       // Shuttle in Place Cnv_Inputs - Need to confirm the order of these Cnv_Inputs.
       // IF (#Cnv_Settings.ID > 110000 AND #Cnv_Settings.ID < 120000 AND NOT #Cnv_Control.Inputs.Sdetect1 AND #Cnv_Control.Inputs.Sdetect2)
       //     OR (#Cnv_Settings.ID > 120000 AND #Cnv_Settings.ID < 130000 AND NOT #Cnv_Control.Inputs.Sdetect1 AND #Cnv_Control.Inputs.Sdetect2) THEN
       //     #Cnv_Control.Error := TRUE; //14:5 Shuttle is about to yeet itself down the VTD shaft
       //     "Set_Bit_F"(Bit := 7,
       //                 Bit_Value := 1,
       //                 Var := #Cnv_Control.Cnv_Errors.Error_Word_2);
       //     #State := 400;
       // END_IF;

       // IF (#Cnv_Settings.ID > 110000 AND #Cnv_Settings.ID < 120000 AND #Cnv_Control.Inputs.Sdetect1 AND NOT #Cnv_Control.Inputs.Sdetect2)
       //     OR (#Cnv_Settings.ID > 120000 AND #Cnv_Settings.ID < 130000 AND #Cnv_Control.Inputs.Sdetect1 AND NOT #Cnv_Control.Inputs.Sdetect2) THEN
       //     #Cnv_Control.Warning := 0; //Shuttle detected in conveyor not yet on barcode
       // END_IF;

       // // #Watchdog auto starts the moment Any form OF transfer occurs.
       // IF #State > 10 AND #State < 400 THEN
       //     #Watchdog(IN := TRUE,
       //               PT := T#200s);
       // ELSE
       //     #Watchdog.IN := FALSE;
       // END_IF;

       // IF #Watchdog.Q THEN
       //     #Watchdog.IN := FALSE;
       //     #Cnv_Control.Error := TRUE; //14:2  Watchdog bit
       //     "Set_Bit_F"(Bit := 4,
       //                 Bit_Value := 1,
       //                 Var := #Cnv_Control.Cnv_Errors.Error_Word_2);
       //     #State := 400;
       // END_IF;

       // go to error state
       IF #Cnv_Control.Cnv_Errors.Error_Word_1 <> 0 OR
           #Cnv_Control.Cnv_Errors.Error_Word_2 <> 0 OR
           #Cnv_Control.Cnv_Errors.Error_Word_3 <> 0 OR
           #Cnv_Control.Cnv_Errors.Error_Word_4 <> 0
       THEN
           #Cnv_Control.Error := TRUE;
           #State := 400;
       END_IF;
   END_REGION

   REGION VFD
       REGION ROLLER
           #Cnv_Control.Roller_Motor.Ready := NOT #Cnv_Control.Roller_Motor.Error;

           #SinaSpeed_Roller(EnableAxis := #Cnv_Control.Roller_Motor.Forward OR #Cnv_Control.Roller_Motor.Reverse,
                             AckError := #Cnv_Control.Instruction.Reset,
                             SpeedSp := #MainSetpoint_Roller,
                             RefSpeed := 1745.0,
                             HWIDSTW := #Cnv_Settings.Roller_G120_Hardware_ID,
                             HWIDZSW := #Cnv_Settings.Roller_G120_Hardware_ID,
                             AxisEnabled => #Cnv_Control.Roller_Motor.Status.%X0,
                             Lockout => #Cnv_Control.Roller_Motor.Error,
                             Error => #Cnv_Control.Roller_Motor.Error);

           //MAIN SETPOINT
           IF #Cnv_Control.Roller_Motor.Reverse THEN
               #MainSetpoint_Roller := (SCALE_X(MIN := 0,
                                                VALUE := NORM_X(MIN := 0,
                                                                VALUE := #Cnv_Control.Roller_Motor.Speed,
                                                                MAX := 100),
                                                MAX := 1745.0) * -1);
           ELSIF #Cnv_Control.Roller_Motor.Forward THEN
               #MainSetpoint_Roller := SCALE_X(MIN := 0,
                                               VALUE := NORM_X(MIN := 0,
                                                               VALUE := #Cnv_Control.Roller_Motor.Speed,
                                                               MAX := 100),
                                               MAX := 1745.0);
           ELSE
               #MainSetpoint_Roller := 0;
           END_IF;

           REGION Actual Speed
               IF #MainSetpoint_Roller > 0 THEN
                   #Cnv_Control.Roller_Motor.Speed_Actual := SCALE_X(MIN := 0,
                                                                     VALUE := NORM_X(MIN := 0,
                                                                                     VALUE := #SinaSpeed_Roller.ActVelocity,
                                                                                     MAX := 1745.0),
                                                                     MAX := 100);
               ELSIF #MainSetpoint_Roller < 0 THEN
                   #Cnv_Control.Roller_Motor.Speed_Actual := SCALE_X(MIN := 0,
                                                                     VALUE := NORM_X(MIN := 0,
                                                                                     VALUE := #SinaSpeed_Roller.ActVelocity * -1,
                                                                                     MAX := 1745.0),
                                                                     MAX := 100);
               ELSE
                   #Cnv_Control.Roller_Motor.Speed_Actual := 0;
               END_IF;
           END_REGION
       END_REGION

       REGION CHAIN
           #Cnv_Control.Chain_Motor.Ready := NOT #Cnv_Control.Chain_Motor.Error;

           #SinaSpeed_Chain(EnableAxis := #Cnv_Control.Chain_Motor.Forward OR #Cnv_Control.Chain_Motor.Reverse,
                            AckError := #Cnv_Control.Instruction.Reset,
                            SpeedSp := #MainSetpoint_Chain,
                            RefSpeed := 1745.0,
                            HWIDSTW := #Cnv_Settings.Chain_G120_Hardware_ID,
                            HWIDZSW := #Cnv_Settings.Chain_G120_Hardware_ID,
                            AxisEnabled => #Cnv_Control.Chain_Motor.Status.%X0,
                            Lockout => #Cnv_Control.Chain_Motor.Error,
                            Error => #Cnv_Control.Chain_Motor.Error);

           //MAIN SETPOINT
           IF #Cnv_Control.Chain_Motor.Reverse THEN
               #MainSetpoint_Chain := (SCALE_X(MIN := 0,
                                               VALUE := NORM_X(MIN := 0,
                                                               VALUE := #Cnv_Control.Chain_Motor.Speed,
                                                               MAX := 100),
                                               MAX := 1745.0) * -1);
           ELSIF #Cnv_Control.Chain_Motor.Forward THEN
               #MainSetpoint_Chain := SCALE_X(MIN := 0,
                                              VALUE := NORM_X(MIN := 0,
                                                              VALUE := #Cnv_Control.Chain_Motor.Speed,
                                                              MAX := 100),
                                              MAX := 1745.0);
           ELSE
               #MainSetpoint_Chain := 0;
           END_IF;

           REGION Actual Speed
               IF #MainSetpoint_Chain > 0 THEN
                   #Cnv_Control.Chain_Motor.Speed_Actual := SCALE_X(MIN := 0,
                                                                    VALUE := NORM_X(MIN := 0,
                                                                                    VALUE := #SinaSpeed_Chain.ActVelocity,
                                                                                    MAX := 1745.0),
                                                                    MAX := 100);
               ELSIF #MainSetpoint_Chain < 0 THEN
                   #Cnv_Control.Chain_Motor.Speed_Actual := SCALE_X(MIN := 0,
                                                                    VALUE := NORM_X(MIN := 0,
                                                                                    VALUE := #SinaSpeed_Chain.ActVelocity * -1,
                                                                                    MAX := 1745.0),
                                                                    MAX := 100);
               ELSE
                   #Cnv_Control.Chain_Motor.Speed_Actual := 0;
               END_IF;
           END_REGION
       END_REGION

       REGION LIFT
           #Cnv_Control.Lift_Motor.Ready := NOT #Cnv_Control.Lift_Motor.Error;

           #SinaSpeed_Lift(EnableAxis := #Cnv_Control.Lift_Motor.Forward OR #Cnv_Control.Lift_Motor.Reverse,
                           AckError := #Cnv_Control.Instruction.Reset,
                           SpeedSp := #MainSetpoint_Lift,
                           RefSpeed := 1745.0,
                           HWIDSTW := #Cnv_Settings.Lift_G120_Hardware_ID,
                           HWIDZSW := #Cnv_Settings.Lift_G120_Hardware_ID,
                           AxisEnabled => #Cnv_Control.Lift_Motor.Status.%X0,
                           Lockout => #Cnv_Control.Lift_Motor.Error,
                           Error => #Cnv_Control.Lift_Motor.Error);

           //MAIN SETPOINT
           IF #Cnv_Control.Lift_Motor.Reverse THEN
               #MainSetpoint_Lift := (SCALE_X(MIN := 0,
                                              VALUE := NORM_X(MIN := 0,
                                                              VALUE := #Cnv_Control.Lift_Motor.Speed,
                                                              MAX := 100),
                                              MAX := 1745.0) * -1);
           ELSIF #Cnv_Control.Lift_Motor.Forward THEN
               #MainSetpoint_Lift := SCALE_X(MIN := 0,
                                             VALUE := NORM_X(MIN := 0,
                                                             VALUE := #Cnv_Control.Lift_Motor.Speed,
                                                             MAX := 100),
                                             MAX := 1745.0);
           ELSE
               #MainSetpoint_Lift := 0;
           END_IF;

           REGION Actual Speed
               IF #MainSetpoint_Lift > 0 THEN
                   #Cnv_Control.Lift_Motor.Speed_Actual := SCALE_X(MIN := 0,
                                                                   VALUE := NORM_X(MIN := 0,
                                                                                   VALUE := #SinaSpeed_Lift.ActVelocity,
                                                                                   MAX := 1745.0),
                                                                   MAX := 100);
               ELSIF #MainSetpoint_Lift < 0 THEN
                   #Cnv_Control.Lift_Motor.Speed_Actual := SCALE_X(MIN := 0,
                                                                   VALUE := NORM_X(MIN := 0,
                                                                                   VALUE := #SinaSpeed_Lift.ActVelocity * -1,
                                                                                   MAX := 1745.0),
                                                                   MAX := 100);
               ELSE
                   #Cnv_Control.Lift_Motor.Speed_Actual := 0;
               END_IF;
           END_REGION
       END_REGION
   END_REGION
END_FUNCTION_BLOCK

FUNCTION_BLOCK "PConveyor_4_FB"   // FB27, SCL
TITLE = Conveyor Instance FB
{ S7_Optimized_Access := 'TRUE' }
AUTHOR : Mertin Coetzee
VERSION : 0.1
// stored: AutoNumber true, IsIECCheckEnabled false, IsRetainMemResEnabled false, MemoryReserve 100, SetENOAutomatically false, UDAEnableTagReadback false
   VAR_INPUT
      Cnv_Settings : "PopUp_Cnv_Settings";
      TimeStartBoost_Roller : UInt;
   END_VAR
   VAR_IN_OUT
      Cnv_Control : "PopUp_Cnv_Control";
      SinaSpeed_Roller : SinaSpeed;
      SinaSpeed_Lift : SinaSpeed;
   END_VAR
   VAR
      State : UInt;
      Timer_TC : TON_TIME;
      Timer_Transfer { S7_SetPoint := 'True'} : TON_TIME;
      Watchdog { S7_SetPoint := 'True'} : TON_TIME;
      Transfer_Direction { S7_SetPoint := 'True'} : String;
      MainSetpoint_Roller : Int;
      MainSetpoint_Lift : Int;
      IEC_Timer_0_Instance_1 { S7_SetPoint := 'True'} : TON_TIME;
      R_TRIG_Instance { S7_SetPoint := 'True'} : R_TRIG;
   END_VAR
   VAR_TEMP
      Execute_Old : Bool;
      Stop_Old : Bool;
   END_VAR
BEGIN
   "R_TRIG_DB_23"(CLK := #Cnv_Control.Instruction.Execute AND NOT #Execute_Old);
   "R_TRIG_DB_24"(CLK := #Cnv_Control.Instruction.Stop AND NOT #Stop_Old);

   #Execute_Old := #Cnv_Control.Instruction.Execute;
   #Stop_Old := #Cnv_Control.Instruction.Stop;

   #Cnv_Control.Enabled := #Cnv_Control.Instruction.Enable;

   //MODES
   #Cnv_Control.Mode := #Cnv_Control.Instruction.Mode_Change;
   IF (#Cnv_Control.Mode = 1 OR #Cnv_Control.Mode = 5) AND NOT #Cnv_Control.Error THEN
       #State := 500;
   END_IF;

   #R_TRIG_Instance(CLK := #Cnv_Control.Mode = 3);
   IF #R_TRIG_Instance.Q THEN
       #State := 0;
   END_IF;

   (*
   TODO:
   01. Need to add statemachine watchdog - Done
   02. Extractor needs to be on same floor for pallet to be moved in manual passed Rbwd - Done
   03. Complete reset state - Done
   04. Add stop inputs - Done
   05. Need to add variable motor speed, manual needs to be slower. - Done
   06. Need to add cyclic error checking. For odd sensor combinations as well - Partially done
   07. Need to add Shuttle monitor - Done
   08. Need to add Task ID check and start bit check to outbound pallet move. Check direction of pallet movement based on connected Cnv.
   09. Need to add checks for wrong direction of travel - Done
   10. Add checks for unsafe conditions with Cnv_Inputs - Partially Done
   11. Define Error codes - DOne
   12. Add watchdof time to Cnv Settings - Done
   13. Add self-timeout on manual 
   14. For shuttle in place sensor checks take into account extractor floor and safety stopper state
   15. Confirm modes and states are correct (Semi-auto and maintenance as well)
   16. Add the correct transfer process for the logistex-spacemaker pallet handovers.

   Mode select is done via the HMI. Might add external mode select switches.

           Mode select mask:
           0: Disabled
           1: Manual
           2: Semi-Auto
           3: Auto
           4: Teach - N/A for Cnv
           5: Maintenance

   Device ID Format: XXYYZZ    
   XX = Device type   
       01   VTD
       10  Cnv_Front_of_VTD
       11  Cnv_Rear_of_VTD
       12  Cnv_On_Extractor
       20  Safety_Stop_Front_of_VTD
       21  Safety_Stop_Rear_of_VTD
   YY = Floor   
   ZZ = VTD Connected to    
   Example: 110203 Conveyor at the rear of VTD 3 on level 2

   Pallet Alignment
   0 = no alignment
   1 = center alignment
   2 = Left
   3 = Right

    Sensor order for the conveyor:
    Lfwd Lpd1 Lpd2
     []   []   []
    ##############################
    #        Pallet Flow         #
    #         ------->>          #
    #                            #
    #                            #
    ##############################
                     []   []   []
                    Rpd2 Rpd1 Rbwd      
   *)


   REGION Cyclic Checks    
       #Cnv_Control.Cnv_Occupied := "PopUp Conveyor 4 - Pallet present 1";

       // Update the Cnv_Control opbject
       #Cnv_Control.SM_State := #State;
       #Cnv_Control.Stopped := NOT #Cnv_Control.Running;
       IF #Cnv_Control.Instruction.Inbound_Ready OR #Cnv_Control.Instruction.Outbound_Ready THEN
           #Cnv_Control.Ready_For_Task := TRUE;
       ELSE
           #Cnv_Control.Ready_For_Task := FALSE;
       END_IF;

   END_REGION

   REGION Auto/Semi auto mode
       CASE #State OF
           0: //IDLE MODE
               #Cnv_Control.Instruction.Transfer_Complete := 0;
               #Cnv_Control.Instruction.Transfer_in_Progress := FALSE;
               #Cnv_Control.Running := FALSE;
               #Cnv_Control.Running := FALSE;
               #Cnv_Control.Roller_Motor.Forward := FALSE;
               #Cnv_Control.Roller_Motor.Reverse := FALSE;
               #Cnv_Control.Roller_Motor.Speed := 0;
               #Cnv_Control.Chain_Motor.Forward := FALSE;
               #Cnv_Control.Chain_Motor.Reverse := FALSE;
               #Cnv_Control.Chain_Motor.Speed := 0;
               #Cnv_Control.Lift_Motor.Forward := FALSE;
               #Cnv_Control.Lift_Motor.Reverse := FALSE;
               #Cnv_Control.Lift_Motor.Speed := 0;
               #Transfer_Direction := '';
               #Timer_Transfer(IN := FALSE,
                               PT := T#0ms);
               "IEC_Timer_0_DB_25".TON(IN := FALSE,
                                       PT := t#0s);
               IF #Cnv_Control.Enabled AND (#Cnv_Control.Mode = 3 OR #Cnv_Control.Mode = 2) AND #Cnv_Control.Error = 0 THEN
                   #State := 10;
               END_IF;

           10: //Standby - Conveyor ready to receive instruction
               IF ("R_TRIG_DB_23".Q OR #Cnv_Control.Instruction.Start_Transfer) THEN
                   //Inbound Transfer
                   IF #Cnv_Control.Instruction.Inbound_Ready AND NOT #Cnv_Control.Running AND #Cnv_Control.Error = 0 THEN
                       IF #Cnv_Control.Inputs."Lift Up" THEN
                           #Cnv_Control.Done := FALSE;
                           #Cnv_Control.Instruction.Transfer_in_Progress := TRUE;
                           #Cnv_Control.Current_Task_ID := #Cnv_Control.Instruction.Task_ID;
                           #State := 20;
                       END_IF;
                       //Outbound Transfer    
                   ELSIF #Cnv_Control.Instruction.Outbound_Ready AND NOT #Cnv_Control.Running AND #Cnv_Control.Error = 0 THEN
                       IF #Cnv_Control.Inputs."Lift Up" THEN
                           #Cnv_Control.Done := FALSE;
                           #Cnv_Control.Instruction.Transfer_in_Progress := TRUE;
                           #Cnv_Control.Current_Task_ID := #Cnv_Control.Instruction.Task_ID;
                           #State := 30;
                       END_IF;
                   END_IF;
               END_IF;

               IF #Cnv_Control.Instruction.Lift_Up THEN
                   #Cnv_Control.Done := FALSE;
                   #State := 60; // Lift UP
               ELSIF #Cnv_Control.Instruction.Lift_Down THEN
                   #Cnv_Control.Done := FALSE;
                   #State := 70; // Lift Down
               END_IF;

           20: // Roller Running (Popup Up)
               #Cnv_Control.Running := TRUE;
               #Cnv_Control.Roller_Motor.Forward := TRUE;
               "IEC_Timer_0_DB_25".TON(IN := TRUE,
                                       PT := UINT_TO_TIME(#TimeStartBoost_Roller) * 1000);

               IF NOT "IEC_Timer_0_DB_25".Q THEN
                   #Cnv_Control.Roller_Motor.Speed := 100.0;
               ELSE
                   #Cnv_Control.Roller_Motor.Speed := #Cnv_Settings.Roller_Full_Speed;
               END_IF;

               #Transfer_Direction := 'Foward';

               IF "R_TRIG_DB_24".Q OR "PopUp Conveyor 4 - Pallet present 1" THEN
                   "IEC_Timer_0_DB_25".TON(IN := FALSE,
                                           PT := t#0s);
                   #Cnv_Control.Done := TRUE;
                   #Cnv_Control.Roller_Motor.Forward := FALSE;
                   #Cnv_Control.Roller_Motor.Reverse := FALSE;
                   #Cnv_Control.Roller_Motor.Speed := 0;
                   #Transfer_Direction := '';
                   #State := 0;
               END_IF;

               //Monitor the transfer progress
               #Timer_Transfer(IN := TRUE,
                               PT := UINT_TO_TIME(#Cnv_Settings.Roller_Transfer_Time) * 1000);
               //If the watchdog bites, kill the process
               IF #Timer_Transfer.Q THEN //14:1 Transfer timed out
                   "Set_Bit_F"(Bit := 3,
                               Bit_Value := 1,
                               Var := #Cnv_Control.Cnv_Errors.Error_Word_2);
               END_IF;

           30: // Roller Running (Popup Up)
               IF "Control_DB".Outbound_Cnv.Motor.Status.%X0 THEN
                   #Cnv_Control.Running := TRUE;
                   #Cnv_Control.Roller_Motor.Forward := TRUE;
                   #Cnv_Control.Roller_Motor.Speed := #Cnv_Settings.Roller_Full_Speed;
                   #Transfer_Direction := 'Foward';
               END_IF;

               IF "R_TRIG_DB_24".Q OR NOT "Outbound Conveyor" THEN
                   #Cnv_Control.Done := TRUE;
                   #Cnv_Control.Roller_Motor.Forward := FALSE;
                   #Cnv_Control.Roller_Motor.Reverse := FALSE;
                   #Cnv_Control.Roller_Motor.Speed := 0;
                   #Transfer_Direction := '';
                   #State := 0;
               END_IF;

               //Monitor the transfer progress
               #Timer_Transfer(IN := TRUE,
                               PT := UINT_TO_TIME(#Cnv_Settings.Roller_Transfer_Time) * 1000);
               //If the watchdog bites, kill the process
               IF #Timer_Transfer.Q THEN //14:1 Transfer timed out
                   "Set_Bit_F"(Bit := 3,
                               Bit_Value := 1,
                               Var := #Cnv_Control.Cnv_Errors.Error_Word_2);
               END_IF;

           60: // Lift Up
               #Cnv_Control.Running := TRUE;
               #Cnv_Control.Lift_Motor.Forward := TRUE;
               #Cnv_Control.Lift_Motor.Speed := #Cnv_Settings.Lift_Full_Speed;
               #Transfer_Direction := 'Up';

               IF #Cnv_Control.Inputs."Lift Up" THEN
                   #Cnv_Control.Done := TRUE;
                   #Cnv_Control.Lift_Motor.Forward := FALSE;
                   #Cnv_Control.Lift_Motor.Reverse := FALSE;
                   #Cnv_Control.Lift_Motor.Speed := 0;
                   #Transfer_Direction := '';
                   #State := 0;
               END_IF;

               //Monitor the transfer progress
               #Timer_Transfer(IN := TRUE,
                               PT := UINT_TO_TIME(#Cnv_Settings.Lift_Transfer_Time) * 1000);
               //If the watchdog bites, kill the process
               IF #Timer_Transfer.Q THEN //14:1 Transfer timed out
                   "Set_Bit_F"(Bit := 3,
                               Bit_Value := 1,
                               Var := #Cnv_Control.Cnv_Errors.Error_Word_2);
               END_IF;

           70: // Lift Down
               #Cnv_Control.Running := TRUE;
               #Cnv_Control.Lift_Motor.Reverse := TRUE;
               #Cnv_Control.Lift_Motor.Speed := #Cnv_Settings.Lift_Full_Speed;
               #Transfer_Direction := 'Down';

               IF #Cnv_Control.Inputs."Lift Down" THEN
                   #Cnv_Control.Done := TRUE;
                   #Cnv_Control.Lift_Motor.Forward := FALSE;
                   #Cnv_Control.Lift_Motor.Reverse := FALSE;
                   #Cnv_Control.Lift_Motor.Speed := 0;
                   #Transfer_Direction := '';
                   #State := 0;
               END_IF;

               //Monitor the transfer progress
               #Timer_Transfer(IN := TRUE,
                               PT := UINT_TO_TIME(#Cnv_Settings.Lift_Transfer_Time) * 1000);
               //If the watchdog bites, kill the process
               IF #Timer_Transfer.Q THEN //14:1 Transfer timed out
                   "Set_Bit_F"(Bit := 3,
                               Bit_Value := 1,
                               Var := #Cnv_Control.Cnv_Errors.Error_Word_2);
               END_IF;

           400: //Error state
               #Cnv_Control.Running := FALSE;
               #Cnv_Control.Roller_Motor.Speed := 0;
               #Cnv_Control.Chain_Motor.Speed := 0;
               #Cnv_Control.Lift_Motor.Speed := 0;
               #Cnv_Control.Roller_Motor.Forward := FALSE;
               #Cnv_Control.Chain_Motor.Forward := FALSE;
               #Cnv_Control.Lift_Motor.Forward := FALSE;
               #Cnv_Control.Roller_Motor.Reverse := FALSE;
               #Cnv_Control.Chain_Motor.Reverse := FALSE;
               #Cnv_Control.Lift_Motor.Reverse := FALSE;
               #Cnv_Control.Instruction.Stop := FALSE;
               #Cnv_Control.Instruction.Transfer_in_Progress := FALSE;
               #Watchdog(IN := FALSE,
                         PT := T#0S);
               #Timer_TC(IN := FALSE,
                         PT := T#0S);
               #Timer_Transfer(IN := FALSE,
                               PT := T#0S);
               #IEC_Timer_0_Instance_1(IN := FALSE,
                                       PT := T#0S);
               IF #Cnv_Control.Instruction.Reset THEN
                   #Cnv_Control.Warning := 0;
                   #Cnv_Control.Current_Task_ID := 0;
                   #Cnv_Control.Error := FALSE; //Reset the conveyor

                   #Cnv_Control.Cnv_Errors.Error_Word_1 := 0;
                   #Cnv_Control.Cnv_Errors.Error_Word_2 := 0;
                   #Cnv_Control.Cnv_Errors.Error_Word_3 := 0;
                   #Cnv_Control.Cnv_Errors.Error_Word_4 := 0;
                   #State := 0;
               END_IF;

           500:
               IF #Cnv_Control.Enabled THEN
                   REGION ROLLER
                       IF #Cnv_Control.Inputs."Lift Up" AND NOT #Cnv_Control.Inputs."Lift Down" THEN
                           IF #Cnv_Control.Instruction.Roller_Fwd OR #Cnv_Control.Instruction.Start_Transfer THEN
                               #Cnv_Control.Roller_Motor.Speed := #Cnv_Settings.Roller_Manual_Speed;
                               #Cnv_Control.Roller_Motor.Forward := TRUE;
                               #Cnv_Control.Running := TRUE;
                           ELSIF #Cnv_Control.Instruction.Roller_Bwd OR #Cnv_Control.Instruction.Start_Transfer_Backward THEN
                               #Cnv_Control.Roller_Motor.Speed := #Cnv_Settings.Roller_Manual_Speed;
                               #Cnv_Control.Roller_Motor.Reverse := TRUE;
                               #Cnv_Control.Running := TRUE;
                           ELSE
                               #Cnv_Control.Roller_Motor.Speed := 0;
                               #Cnv_Control.Roller_Motor.Forward := FALSE;
                               #Cnv_Control.Roller_Motor.Reverse := FALSE;
                               #Cnv_Control.Running := FALSE;
                           END_IF;
                       END_IF;
                   END_REGION

                   REGION LIFT
                       IF NOT #SinaSpeed_Roller.AxisEnabled THEN
                           IF #Cnv_Control.Instruction.Lift_Up AND NOT #Cnv_Control.Inputs."Lift Up" THEN
                               #Cnv_Control.Lift_Motor.Speed := #Cnv_Settings.Lift_Manual_Speed;
                               #Cnv_Control.Lift_Motor.Forward := TRUE;
                               #Cnv_Control.Running := TRUE;
                           ELSIF #Cnv_Control.Instruction.Lift_Down AND NOT #Cnv_Control.Inputs."Lift Down" THEN
                               #Cnv_Control.Lift_Motor.Speed := #Cnv_Settings.Lift_Manual_Speed;
                               #Cnv_Control.Lift_Motor.Reverse := TRUE;
                               #Cnv_Control.Running := TRUE;
                           ELSE
                               #Cnv_Control.Lift_Motor.Speed := 0;
                               #Cnv_Control.Lift_Motor.Forward := FALSE;
                               #Cnv_Control.Lift_Motor.Reverse := FALSE;
                               #Cnv_Control.Running := FALSE;
                           END_IF;
                       END_IF;
                   END_REGION
               END_IF;

               IF #Cnv_Control.Mode <> 1 AND #Cnv_Control.Mode <> 5 THEN
                   #State := 0;
               END_IF;
       END_CASE;
   END_REGION



   REGION Cyclic Error Checks
       IF NOT "Main_Safety_RTG1_DB".SAFETY_OK_CAROUSEL THEN //11:1
           "Set_Bit_F"(Bit := 0,
                       Bit_Value := 1,
                       Var := #Cnv_Control.Cnv_Errors.Error_Word_1);
       END_IF;

       // IF #Cnv_Control.Instruction.Stop THEN //11:2
       //     "Set_Bit_F"(Bit := 1,
       //                 Bit_Value := 1,
       //                 Var := #Cnv_Control.Cnv_Errors.Error_Word_1);
       // END_IF;

       IF #Cnv_Control.Roller_Motor.Error OR #Cnv_Control.Chain_Motor.Error OR #Cnv_Control.Lift_Motor.Error THEN
           "Set_Bit_F"(Bit := 0,
                       Bit_Value := 1,
                       Var := #Cnv_Control.Cnv_Errors.Error_Word_4);
       END_IF;

       // Pallet Sensor Checks
       // IF #Cnv_Control.Inputs.Lfwd AND #Cnv_Control.Inputs.Rbwd THEN
       //     #Cnv_Control.Error := TRUE; //15:2 Combination of Cnv_Inputs indicates issue in conveyor
       //     "Set_Bit_F"(Bit := 1,
       //                 Bit_Value := 1,
       //                 Var := #Cnv_Control.Cnv_Errors.Error_Word_4);
       //     #State := 400;
       // IF #Cnv_Control.Inputs.Lfwd AND #Cnv_Control.Inputs.Lpd1 AND #Cnv_Control.Inputs.Rpd1 THEN
       //     #Cnv_Control.Error := TRUE; //15:3 Combination of Cnv_Inputs indicates issue in conveyor
       //     "Set_Bit_F"(Bit := 2,
       //                 Bit_Value := 1,
       //                 Var := #Cnv_Control.Cnv_Errors.Error_Word_4);
       //     #State := 400;
       // ELSIF #Cnv_Control.Inputs.Rbwd AND #Cnv_Control.Inputs.Lpd1 AND #Cnv_Control.Inputs.Rpd1 THEN
       //     #Cnv_Control.Error := TRUE; //15:4 Combination of Cnv_Inputs indicates issue in conveyor
       //     "Set_Bit_F"(Bit := 3,
       //                 Bit_Value := 1,
       //                 Var := #Cnv_Control.Cnv_Errors.Error_Word_4);
       //     #State := 400;
       // END_IF;

       // Shuttle in Place Cnv_Inputs - Need to confirm the order of these Cnv_Inputs.
       // IF (#Cnv_Settings.ID > 110000 AND #Cnv_Settings.ID < 120000 AND NOT #Cnv_Control.Inputs.Sdetect1 AND #Cnv_Control.Inputs.Sdetect2)
       //     OR (#Cnv_Settings.ID > 120000 AND #Cnv_Settings.ID < 130000 AND NOT #Cnv_Control.Inputs.Sdetect1 AND #Cnv_Control.Inputs.Sdetect2) THEN
       //     #Cnv_Control.Error := TRUE; //14:5 Shuttle is about to yeet itself down the VTD shaft
       //     "Set_Bit_F"(Bit := 7,
       //                 Bit_Value := 1,
       //                 Var := #Cnv_Control.Cnv_Errors.Error_Word_2);
       //     #State := 400;
       // END_IF;

       // IF (#Cnv_Settings.ID > 110000 AND #Cnv_Settings.ID < 120000 AND #Cnv_Control.Inputs.Sdetect1 AND NOT #Cnv_Control.Inputs.Sdetect2)
       //     OR (#Cnv_Settings.ID > 120000 AND #Cnv_Settings.ID < 130000 AND #Cnv_Control.Inputs.Sdetect1 AND NOT #Cnv_Control.Inputs.Sdetect2) THEN
       //     #Cnv_Control.Warning := 0; //Shuttle detected in conveyor not yet on barcode
       // END_IF;

       // // #Watchdog auto starts the moment Any form OF transfer occurs.
       // IF #State > 10 AND #State < 400 THEN
       //     #Watchdog(IN := TRUE,
       //               PT := T#200s);
       // ELSE
       //     #Watchdog.IN := FALSE;
       // END_IF;

       // IF #Watchdog.Q THEN
       //     #Watchdog.IN := FALSE;
       //     #Cnv_Control.Error := TRUE; //14:2  Watchdog bit
       //     "Set_Bit_F"(Bit := 4,
       //                 Bit_Value := 1,
       //                 Var := #Cnv_Control.Cnv_Errors.Error_Word_2);
       //     #State := 400;
       // END_IF;

       // go to error state
       IF #Cnv_Control.Cnv_Errors.Error_Word_1 <> 0 OR
           #Cnv_Control.Cnv_Errors.Error_Word_2 <> 0 OR
           #Cnv_Control.Cnv_Errors.Error_Word_3 <> 0 OR
           #Cnv_Control.Cnv_Errors.Error_Word_4 <> 0
       THEN
           #Cnv_Control.Error := TRUE;
           #State := 400;
       END_IF;
   END_REGION

   REGION VFD
       REGION ROLLER
           #Cnv_Control.Roller_Motor.Ready := NOT #Cnv_Control.Roller_Motor.Error;

           #SinaSpeed_Roller(EnableAxis := #Cnv_Control.Roller_Motor.Forward OR #Cnv_Control.Roller_Motor.Reverse,
                             AckError := #Cnv_Control.Instruction.Reset,
                             SpeedSp := #MainSetpoint_Roller,
                             RefSpeed := 1745.0,
                             HWIDSTW := #Cnv_Settings.Roller_G120_Hardware_ID,
                             HWIDZSW := #Cnv_Settings.Roller_G120_Hardware_ID,
                             AxisEnabled => #Cnv_Control.Roller_Motor.Status.%X0,
                             Lockout => #Cnv_Control.Roller_Motor.Error,
                             Error => #Cnv_Control.Roller_Motor.Error);

           //MAIN SETPOINT
           IF #Cnv_Control.Roller_Motor.Reverse THEN
               #MainSetpoint_Roller := (SCALE_X(MIN := 0,
                                                VALUE := NORM_X(MIN := 0,
                                                                VALUE := #Cnv_Control.Roller_Motor.Speed,
                                                                MAX := 100),
                                                MAX := 1745.0) * -1);
           ELSIF #Cnv_Control.Roller_Motor.Forward THEN
               #MainSetpoint_Roller := SCALE_X(MIN := 0,
                                               VALUE := NORM_X(MIN := 0,
                                                               VALUE := #Cnv_Control.Roller_Motor.Speed,
                                                               MAX := 100),
                                               MAX := 1745.0);
           ELSE
               #MainSetpoint_Roller := 0;
           END_IF;

           REGION Actual Speed
               IF #MainSetpoint_Roller > 0 THEN
                   #Cnv_Control.Roller_Motor.Speed_Actual := SCALE_X(MIN := 0,
                                                                     VALUE := NORM_X(MIN := 0,
                                                                                     VALUE := #SinaSpeed_Roller.ActVelocity,
                                                                                     MAX := 1745.0),
                                                                     MAX := 100);
               ELSIF #MainSetpoint_Roller < 0 THEN
                   #Cnv_Control.Roller_Motor.Speed_Actual := SCALE_X(MIN := 0,
                                                                     VALUE := NORM_X(MIN := 0,
                                                                                     VALUE := #SinaSpeed_Roller.ActVelocity * -1,
                                                                                     MAX := 1745.0),
                                                                     MAX := 100);
               ELSE
                   #Cnv_Control.Roller_Motor.Speed_Actual := 0;
               END_IF;
           END_REGION
       END_REGION

       REGION LIFT
           #Cnv_Control.Lift_Motor.Ready := NOT #Cnv_Control.Lift_Motor.Error;

           #SinaSpeed_Lift(EnableAxis := #Cnv_Control.Lift_Motor.Forward OR #Cnv_Control.Lift_Motor.Reverse,
                           AckError := #Cnv_Control.Instruction.Reset,
                           SpeedSp := #MainSetpoint_Lift,
                           RefSpeed := 1745.0,
                           HWIDSTW := #Cnv_Settings.Lift_G120_Hardware_ID,
                           HWIDZSW := #Cnv_Settings.Lift_G120_Hardware_ID,
                           AxisEnabled => #Cnv_Control.Lift_Motor.Status.%X0,
                           Lockout => #Cnv_Control.Lift_Motor.Error,
                           Error => #Cnv_Control.Lift_Motor.Error);

           //MAIN SETPOINT
           IF #Cnv_Control.Lift_Motor.Reverse THEN
               #MainSetpoint_Lift := (SCALE_X(MIN := 0,
                                              VALUE := NORM_X(MIN := 0,
                                                              VALUE := #Cnv_Control.Lift_Motor.Speed,
                                                              MAX := 100),
                                              MAX := 1745.0) * -1);
           ELSIF #Cnv_Control.Lift_Motor.Forward THEN
               #MainSetpoint_Lift := SCALE_X(MIN := 0,
                                             VALUE := NORM_X(MIN := 0,
                                                             VALUE := #Cnv_Control.Lift_Motor.Speed,
                                                             MAX := 100),
                                             MAX := 1745.0);
           ELSE
               #MainSetpoint_Lift := 0;
           END_IF;

           REGION Actual Speed
               IF #MainSetpoint_Lift > 0 THEN
                   #Cnv_Control.Lift_Motor.Speed_Actual := SCALE_X(MIN := 0,
                                                                   VALUE := NORM_X(MIN := 0,
                                                                                   VALUE := #SinaSpeed_Lift.ActVelocity,
                                                                                   MAX := 1745.0),
                                                                   MAX := 100);
               ELSIF #MainSetpoint_Lift < 0 THEN
                   #Cnv_Control.Lift_Motor.Speed_Actual := SCALE_X(MIN := 0,
                                                                   VALUE := NORM_X(MIN := 0,
                                                                                   VALUE := #SinaSpeed_Lift.ActVelocity * -1,
                                                                                   MAX := 1745.0),
                                                                   MAX := 100);
               ELSE
                   #Cnv_Control.Lift_Motor.Speed_Actual := 0;
               END_IF;
           END_REGION
       END_REGION
   END_REGION
END_FUNCTION_BLOCK

FUNCTION_BLOCK "PickConveyor_FB"   // FB35, SCL
TITLE = Conveyor Instance FB
{ S7_Optimized_Access := 'TRUE' }
AUTHOR : Mertin Coetzee
VERSION : 0.1
// stored: AutoNumber true, IsIECCheckEnabled false, IsRetainMemResEnabled false, MemoryReserve 100, SetENOAutomatically false, UDAEnableTagReadback false
   VAR_INPUT
      Cnv_Settings : "Pick_Cnv_Settings";
   END_VAR
   VAR_IN_OUT
      SinaSpeed_Chain : SinaSpeed;
   END_VAR
   VAR
      State : UInt;
      Timer_TC : TON_TIME;
      Timer_Transfer { S7_SetPoint := 'True'} : TON_TIME;
      Watchdog { S7_SetPoint := 'True'} : TON_TIME;
      Transfer_Direction { S7_SetPoint := 'True'} : String;
      MainSetpoint_Chain : Int;
      IEC_Timer_0_Instance_1 { S7_SetPoint := 'True'} : TON_TIME;
      R_TRIG_Instance { S7_SetPoint := 'True'} : R_TRIG;
   END_VAR
   VAR_TEMP
      Execute_Old : Bool;
      Stop_Old : Bool;
   END_VAR
BEGIN
   "R_TRIG_DB_28"(CLK := "Control_DB".Pick_Station.Instruction.Execute AND NOT #Execute_Old);
   "R_TRIG_DB_29"(CLK := "Control_DB".Pick_Station.Instruction.Stop AND NOT #Stop_Old);

   #Execute_Old := "Control_DB".Pick_Station.Instruction.Execute;
   #Stop_Old := "Control_DB".Pick_Station.Instruction.Stop;

   "Control_DB".Pick_Station.Enabled := "Control_DB".Pick_Station.Instruction.Enable;

   //MODES
   "Control_DB".Pick_Station.Mode := "Control_DB".Pick_Station.Instruction.Mode_Change;
   IF ("Control_DB".Pick_Station.Mode = 1 OR "Control_DB".Pick_Station.Mode = 5) AND NOT "Control_DB".Pick_Station.Error THEN
       #State := 500;
   END_IF;

   #R_TRIG_Instance(CLK := "Control_DB".Pick_Station.Mode = 3);
   IF #R_TRIG_Instance.Q THEN
       #State := 0;
   END_IF;

   (*
   TODO:
   01. Need to add statemachine watchdog - Done
   02. Extractor needs to be on same floor for pallet to be moved in manual passed Rbwd - Done
   03. Complete reset state - Done
   04. Add stop inputs - Done
   05. Need to add variable motor speed, manual needs to be slower. - Done
   06. Need to add cyclic error checking. For odd sensor combinations as well - Partially done
   07. Need to add Shuttle monitor - Done
   08. Need to add Task ID check and start bit check to outbound pallet move. Check direction of pallet movement based on connected Cnv.
   09. Need to add checks for wrong direction of travel - Done
   10. Add checks for unsafe conditions with Cnv_Inputs - Partially Done
   11. Define Error codes - DOne
   12. Add watchdof time to Cnv Settings - Done
   13. Add self-timeout on manual 
   14. For shuttle in place sensor checks take into account extractor floor and safety stopper state
   15. Confirm modes and states are correct (Semi-auto and maintenance as well)
   16. Add the correct transfer process for the logistex-spacemaker pallet handovers.

   Mode select is done via the HMI. Might add external mode select switches.

           Mode select mask:
           0: Disabled
           1: Manual
           2: Semi-Auto
           3: Auto
           4: Teach - N/A for Cnv
           5: Maintenance

   Device ID Format: XXYYZZ    
   XX = Device type   
       01   VTD
       10  Cnv_Front_of_VTD
       11  Cnv_Rear_of_VTD
       12  Cnv_On_Extractor
       20  Safety_Stop_Front_of_VTD
       21  Safety_Stop_Rear_of_VTD
   YY = Floor   
   ZZ = VTD Connected to    
   Example: 110203 Conveyor at the rear of VTD 3 on level 2

   Pallet Alignment
   0 = no alignment
   1 = center alignment
   2 = Left
   3 = Right

    Sensor order for the conveyor:
    Lfwd Lpd1 Lpd2
     []   []   []
    ##############################
    #        Pallet Flow         #
    #         ------->>          #
    #                            #
    #                            #
    ##############################
                     []   []   []
                    Rpd2 Rpd1 Rbwd      
   *)

   REGION Cyclic Checks    
       // Update the pallet type as the Cnv_Inputs are triggered.
       "Control_DB".Pick_Station.Cnv_Occupied := NOT "Pick Station";

       // Update the Cnv_Control opbject
       "Control_DB".Pick_Station.SM_State := #State;
       "Control_DB".Pick_Station.Stopped := NOT "Control_DB".Pick_Station.Running;
       IF "Control_DB".Pick_Station.Instruction.Inbound_Ready OR "Control_DB".Pick_Station.Instruction.Outbound_Ready THEN
           "Control_DB".Pick_Station.Ready_For_Task := TRUE;
       ELSE
           "Control_DB".Pick_Station.Ready_For_Task := FALSE;
       END_IF;
   END_REGION

   REGION Auto/Semi auto mode
       CASE #State OF
           0: //Initialization
               "Control_DB".Pick_Station.Instruction.Transfer_Complete := 0;
               "Control_DB".Pick_Station.Instruction.Transfer_in_Progress := FALSE;
               "Control_DB".Pick_Station.Running := FALSE;
               "Control_DB".Pick_Station.Motor.Forward := FALSE;
               "Control_DB".Pick_Station.Motor.Reverse := FALSE;
               "Control_DB".Pick_Station.Motor.Speed := 0;
               #Transfer_Direction := '';
               #Timer_Transfer(IN := FALSE,
                               PT := T#0ms);
               IF "Control_DB".Pick_Station.Enabled AND ("Control_DB".Pick_Station.Mode = 3 OR "Control_DB".Pick_Station.Mode = 2) AND "Control_DB".Pick_Station.Error = 0 THEN
                   #State := 10;
               END_IF;

           10: //Standby - Conveyor ready to receive instruction
               IF ("R_TRIG_DB_28".Q OR "Control_DB".Pick_Station.Instruction.Start_Transfer) THEN
                   //Inbound Transfer
                   IF "Control_DB".Pick_Station.Instruction.Inbound_Ready AND NOT "Control_DB".Pick_Station.Running AND "Control_DB".Pick_Station.Error = 0 THEN
                       //Check sensors
                       IF "Control_DB".PopUp_Cnv[4].Inputs."Lift Down" THEN //TO pick station
                           "Control_DB".Pick_Station.Done := FALSE;
                           "Control_DB".Pick_Station.Instruction.Transfer_in_Progress := TRUE;
                           "Control_DB".Pick_Station.Current_Task_ID := "Control_DB".Pick_Station.Instruction.Task_ID;
                           #State := 30;// Chain Running (Popup Down) 
                       ELSE
                           "Control_DB".Pick_Station.Warning := 1; //Cannot transfer from that conveyor
                       END_IF;

                       //Outbound Transfer    
                   ELSIF "Control_DB".Pick_Station.Instruction.Outbound_Ready AND NOT "Control_DB".Pick_Station.Running AND "Control_DB".Pick_Station.Error = 0 THEN
                       //Check sensors
                       IF "Control_DB".PopUp_Cnv[1].Inputs."Lift Down"  THEN
                           "Control_DB".Pick_Station.Done := FALSE;
                           "Control_DB".Pick_Station.Instruction.Transfer_in_Progress := TRUE;
                           "Control_DB".Pick_Station.Current_Task_ID := "Control_DB".Pick_Station.Instruction.Task_ID;
                           #State := 40;
                       ELSE
                           "Control_DB".Pick_Station.Warning := 1; //Cannot transfer TO that conveyor
                       END_IF;
                   ELSE
                       "Control_DB".Pick_Station.Warning := 0;// No task that can be started, yet start bit has been made true.
                   END_IF;
               ELSIF "Control_DB".Pick_Station.Instruction.Start_Transfer AND "Control_DB".VTD_Control.Current_Level <> 0 THEN
                   //Extractor not at the correct level
                   "Set_Bit_F"(Bit := 2,
                               Bit_Value := 1,
                               Var := "Control_DB".Pick_Station.Cnv_Errors.Error_Word_3);
               END_IF;

           30: // Chain Running (Popup Down)
               "Control_DB".Pick_Station.Running := TRUE;
               "Control_DB".Pick_Station.Motor.Forward := TRUE;
               "Control_DB".Pick_Station.Motor.Speed := #Cnv_Settings.Full_Speed;
               #Transfer_Direction := 'Foward';

               IF "R_TRIG_DB_29".Q OR NOT "Pick Station" THEN
                   "Control_DB".Pick_Station.Done := TRUE;
                   "Control_DB".Pick_Station.Motor.Forward := FALSE;
                   "Control_DB".Pick_Station.Motor.Reverse := FALSE;
                   "Control_DB".Pick_Station.Motor.Speed := 0;
                   #Transfer_Direction := '';
                   #State := 0;
               END_IF;

               //Monitor the transfer progress
               #Timer_Transfer(IN := "IEC_Timer_0_DB_21".Q,
                               PT := UINT_TO_TIME(#Cnv_Settings.Transfer_Time) * 1000);
               //If the watchdog bites, kill the process
               IF #Timer_Transfer.Q THEN //14:1 Transfer timed out
                   "Set_Bit_F"(Bit := 3,
                               Bit_Value := 1,
                               Var := "Control_DB".Pick_Station.Cnv_Errors.Error_Word_2);
               END_IF;

           40: // Chain Running (Popup Down)
               "Control_DB".Pick_Station.Running := TRUE;
               "Control_DB".Pick_Station.Motor.Forward := TRUE;
               "Control_DB".Pick_Station.Motor.Speed := #Cnv_Settings.Full_Speed;
               #Transfer_Direction := 'Foward';

               IF "R_TRIG_DB_29".Q OR "PopUp Conveyor 1 - Pallet sensor" THEN
                   "Control_DB".Pick_Station.Done := TRUE;
                   "Control_DB".Pick_Station.Motor.Forward := FALSE;
                   "Control_DB".Pick_Station.Motor.Reverse := FALSE;
                   "Control_DB".Pick_Station.Motor.Speed := 0;
                   #Transfer_Direction := '';
                   #State := 0;
               END_IF;

               //Monitor the transfer progress
               #Timer_Transfer(IN := "IEC_Timer_0_DB_21".Q,
                               PT := UINT_TO_TIME(#Cnv_Settings.Transfer_Time) * 1000);
               //If the watchdog bites, kill the process
               IF #Timer_Transfer.Q THEN //14:1 Transfer timed out
                   "Set_Bit_F"(Bit := 3,
                               Bit_Value := 1,
                               Var := "Control_DB".Pick_Station.Cnv_Errors.Error_Word_2);
               END_IF;

           400: //Error state
               "Control_DB".Pick_Station.Running := FALSE;
               "Control_DB".Pick_Station.Motor.Speed := 0;
               "Control_DB".Pick_Station.Motor.Forward := FALSE;
               "Control_DB".Pick_Station.Motor.Reverse := FALSE;
               "Control_DB".Pick_Station.Instruction.Stop := FALSE;
               "Control_DB".Pick_Station.Instruction.Transfer_in_Progress := FALSE;
               #Watchdog(IN := FALSE,
                         PT := T#0S);
               #Timer_TC(IN := FALSE,
                         PT := T#0S);
               #Timer_Transfer(IN := FALSE,
                               PT := T#0S);
               #IEC_Timer_0_Instance_1(IN := FALSE,
                                       PT := T#0S);
               IF "Control_DB".Pick_Station.Instruction.Reset THEN
                   "Control_DB".Pick_Station.Warning := 0;
                   "Control_DB".Pick_Station.Current_Task_ID := 0;
                   "Control_DB".Pick_Station.Error := FALSE; //Reset the conveyor

                   "Control_DB".Pick_Station.Cnv_Errors.Error_Word_1 := 0;
                   "Control_DB".Pick_Station.Cnv_Errors.Error_Word_2 := 0;
                   "Control_DB".Pick_Station.Cnv_Errors.Error_Word_3 := 0;
                   "Control_DB".Pick_Station.Cnv_Errors.Error_Word_4 := 0;
                   #State := 0;
               END_IF;

           500:
               IF "Control_DB".Pick_Station.Enabled THEN
                   IF "Control_DB".Pick_Station.Instruction.Foward OR "Control_DB".Pick_Station.Instruction.Start_Transfer THEN
                       "Control_DB".Pick_Station.Motor.Speed := #Cnv_Settings.Manual_Speed;
                       "Control_DB".Pick_Station.Motor.Forward := TRUE;
                       "Control_DB".Pick_Station.Running := TRUE;
                   ELSIF "Control_DB".Pick_Station.Instruction.Backward OR "Control_DB".Pick_Station.Instruction.Start_Transfer_Backward THEN
                       "Control_DB".Pick_Station.Motor.Speed := #Cnv_Settings.Manual_Speed;
                       "Control_DB".Pick_Station.Motor.Reverse := TRUE;
                       "Control_DB".Pick_Station.Running := TRUE;
                   ELSE
                       "Control_DB".Pick_Station.Motor.Speed := 0;
                       "Control_DB".Pick_Station.Motor.Forward := FALSE;
                       "Control_DB".Pick_Station.Motor.Reverse := FALSE;
                       "Control_DB".Pick_Station.Running := FALSE;
                   END_IF;
               END_IF;

               IF "Control_DB".Pick_Station.Mode <> 1 AND "Control_DB".Pick_Station.Mode <> 5 THEN
                   #State := 0;
               END_IF;
       END_CASE;
   END_REGION



   REGION Cyclic Error Checks
       IF NOT "Main_Safety_RTG1_DB".SAFETY_OK_CAROUSEL THEN //11:1
           "Set_Bit_F"(Bit := 0,
                       Bit_Value := 1,
                       Var := "Control_DB".Pick_Station.Cnv_Errors.Error_Word_1);
       END_IF;

       IF "Control_DB".Pick_Station.Motor.Error THEN
           "Set_Bit_F"(Bit := 0,
                       Bit_Value := 1,
                       Var := "Control_DB".Pick_Station.Cnv_Errors.Error_Word_4);
       END_IF;

       // go to error state
       IF "Control_DB".Pick_Station.Cnv_Errors.Error_Word_1 <> 0 OR
           "Control_DB".Pick_Station.Cnv_Errors.Error_Word_2 <> 0 OR
           "Control_DB".Pick_Station.Cnv_Errors.Error_Word_3 <> 0 OR
           "Control_DB".Pick_Station.Cnv_Errors.Error_Word_4 <> 0
       THEN
           "Control_DB".Pick_Station.Error := TRUE;
           #State := 400;
       END_IF;
   END_REGION

   REGION VFD
       "IEC_Timer_0_DB_21".TON(IN:="LighGuard_Cut-Off Path 01",
                               PT:=T#3s);

       "Control_DB".Pick_Station.Motor.Ready := NOT "Control_DB".Pick_Station.Motor.Error;

       #SinaSpeed_Chain(EnableAxis := ("Control_DB".Pick_Station.Motor.Forward OR "Control_DB".Pick_Station.Motor.Reverse) AND "IEC_Timer_0_DB_21".Q,
                        AckError := "Control_DB".Pick_Station.Instruction.Reset,
                            SpeedSp := #MainSetpoint_Chain,
                            RefSpeed := 1745.0,
                            HWIDSTW := #Cnv_Settings.G120_Hardware_ID,
                            HWIDZSW := #Cnv_Settings.G120_Hardware_ID,
                            AxisEnabled => "Control_DB".Pick_Station.Motor.Status.%X0,
                            Lockout => "Control_DB".Pick_Station.Motor.Error,
                            Error => "Control_DB".Pick_Station.Motor.Error);

           //MAIN SETPOINT
           IF "Control_DB".Pick_Station.Motor.Reverse AND "IEC_Timer_0_DB_21".Q THEN
               #MainSetpoint_Chain := (SCALE_X(MIN := 0,
                                               VALUE := NORM_X(MIN := 0,
                                                               VALUE := "Control_DB".Pick_Station.Motor.Speed,
                                                               MAX := 100),
                                               MAX := 1745.0) * -1);
           ELSIF "Control_DB".Pick_Station.Motor.Forward AND "IEC_Timer_0_DB_21".Q THEN
               #MainSetpoint_Chain := SCALE_X(MIN := 0,
                                              VALUE := NORM_X(MIN := 0,
                                                              VALUE := "Control_DB".Pick_Station.Motor.Speed,
                                                              MAX := 100),
                                              MAX := 1745.0);
           ELSE
               #MainSetpoint_Chain := 0;
           END_IF;

           REGION Actual Speed
               IF #MainSetpoint_Chain > 0 THEN
                   "Control_DB".Pick_Station.Motor.Speed_Actual := SCALE_X(MIN := 0,
                                                                    VALUE := NORM_X(MIN := 0,
                                                                                    VALUE := #SinaSpeed_Chain.ActVelocity,
                                                                                    MAX := 1745.0),
                                                                    MAX := 100);
               ELSIF #MainSetpoint_Chain < 0 THEN
                   "Control_DB".Pick_Station.Motor.Speed_Actual := SCALE_X(MIN := 0,
                                                                    VALUE := NORM_X(MIN := 0,
                                                                                    VALUE := #SinaSpeed_Chain.ActVelocity * -1,
                                                                                    MAX := 1745.0),
                                                                    MAX := 100);
               ELSE
                   "Control_DB".Pick_Station.Motor.Speed_Actual := 0;
               END_IF;
           END_REGION
    END_REGION
END_FUNCTION_BLOCK

FUNCTION_BLOCK "VTD_FB"   // FB18, SCL
{ S7_Optimized_Access := 'TRUE' }
VERSION : 0.1
// stored: AutoNumber true, IsIECCheckEnabled false, IsRetainMemResEnabled false, MemoryReserve 100, SetENOAutomatically false, UDAEnableTagReadback false
   VAR_INPUT
      Cnv_Sensors : "ECnv_Inputs";
      VTD_Settings : "VTD_Settings";
   END_VAR
   VAR_IN_OUT
      VTD_Control : "VTD_Control";
      SinaSpeed : SinaSpeed;
   END_VAR
   VAR
      State : UInt;
      I_State : UInt;
      LD_Timer : TON_TIME;
      LP_Timer { S7_SetPoint := 'True'} : TON_TIME;
      Watchdog { S7_SetPoint := 'True'} : TON_TIME;
      CS_TImer { S7_SetPoint := 'True'} : TON_TIME;
      Interlock_Timer { S7_SetPoint := 'True'} : TON_TIME;
      MainSetpoint : Int;
      Position_Offset : Real;
      ChangeToLow : Array[1..4] of DInt;
      DestPosition : Real;
      SetUpSpeed : UInt;
      LevelBelowExtractor : UInt := 1;
      IEC_Timer_0_Instance { S7_SetPoint := 'True'} : TON_TIME;
      DestinationLevel : UInt;
      CurrentlLevel : UInt;
      VTD_ID_Decoded { ExternalAccessible := 'False'; ExternalVisible := 'False'; ExternalWritable := 'False'} : "ID_Decoded";
      Cnv_ID_Decoded { ExternalAccessible := 'False'; ExternalVisible := 'False'; ExternalWritable := 'False'} : "ID_Decoded";
      IEC_Timer_0_Instance_1 { S7_SetPoint := 'True'} : TON_TIME;
      IEC_Timer_0_Instance_2 { S7_SetPoint := 'True'} : TON_TIME;
      VTD_ControlInstructionTask_ID_Old : Int;
      R_Execulte { S7_SetPoint := 'True'} : R_TRIG;
   END_VAR
   VAR_TEMP
      Level_Accuracy : String;
      i : UInt;
      Do_Once : Bool;
      Level_Detect : Bool;
      Upper_limit : Bool;
      Lower_Limit : Bool;
      Ultimate_Slow : Bool;
      Ulitmate_Creep : Bool;
      Level_Detect2 : Bool;
      Level_Detect1 : Bool;
      LPR_Extended : Bool;
      LPR_Retracted : Bool;
      LPL_Extended : Bool;
      LPL_Retracted : Bool;
      Shuttle_Detect1 : Bool;
      Shuttle_Detect2 : Bool;
      LPL_Retract : Bool;
      LPL_Extend : Bool;
      LPR_Retract : Bool;
      LPR_Extend : Bool;
      Cnvs1_NotExtended : Bool;
      Cnvs2_NotExtended : Bool;
      Stoppers_NotExtended : Bool;
      MainSetpoint1 : Int;
   END_VAR
BEGIN
   //Execute
   #R_Execulte(CLK:=#VTD_Control.Instruction.Execulte);

   IF #VTD_Control.Mode = 3 THEN
       #VTD_Control.Instruction.Enable := TRUE;
   END_IF;

   #VTD_Control.Enabled := #VTD_Control.Instruction.Enable;

   #VTD_Control.Mode := "Control_DB".VTD_Control.Instruction.Mode_Change;

   //MANUAL MODE
   IF (#VTD_Control.Mode = 1 OR #VTD_Control.Mode = 5) AND NOT #VTD_Control.Error THEN
       #State := 500;
   END_IF;

   (*
   TODO:

   Mode select is done via the HMI. Might add external mode select switches.

           Mode select mask:
           0: Disabled
           1: Manual
           2: Semi-Auto
           3: Auto
           4: Teach
           5: Maintenance

   Device ID Format: XXYYZZ    
   XX = Device type   
       01   VTD
       10  Cnv_Front_of_VTD
       11  Cnv_Rear_of_VTD
       12  Cnv_On_Extractor
       20  Safety_Stop_Front_of_VTD
       21  Safety_Stop_Rear_of_VTD
   YY = Floor   
   ZZ = VTD Connected to 
   *)

   REGION Sensor allocations
       //Assign inputs to local vars
       #Upper_limit := "Upper Ultimate";
       #Lower_Limit := "Lower Ultimate";
       #Ultimate_Slow := "Slowdown";
       #Ulitmate_Creep := "Creep speed";
       #Level_Detect2 := "Docking Sensor Rear";
       #Level_Detect1 := "Docking Sensor Front";
       #LPR_Extended := "Locking Pins Extended Right";
       #LPR_Retracted := "Locking Pins Retracted Right";
       #LPL_Extended := "Locking Pins Extended left";
       #LPL_Retracted := "Locking Pins Retracted left";

       #VTD_Control.LE := "LE_X_Unsafe_Position_1";
       #VTD_Control.AE := "AE_Position_1_Scaled";
   END_REGION

   REGION Cyclic Checks
       // Check for shuttle
       IF #Shuttle_Detect1 AND #Shuttle_Detect2 THEN
           #VTD_Control.Shuttle_Loaded := 1; //inplace
       ELSIF NOT #Shuttle_Detect1 AND #Shuttle_Detect2 THEN
           #VTD_Control.Shuttle_Loaded := 2; // Front overhang
       ELSIF #Shuttle_Detect1 AND NOT #Shuttle_Detect2 THEN
           #VTD_Control.Shuttle_Loaded := 3; //Rear overhang
       ELSE
           #VTD_Control.Shuttle_Loaded := 0; //None
       END_IF;

       // Check for Pallet
       IF #Cnv_Sensors."Pallet Detect 1" OR #Cnv_Sensors."Pallet Detect 2" THEN
           //Chep Pallet
           IF #Cnv_Sensors."Pallet Detect 1" AND #Cnv_Sensors."Pallet Detect 2" THEN
               #VTD_Control.Pallet_Loaded := 2; //Chep
               //Euro skewed to the left
           ELSIF #Cnv_Sensors."Pallet Detect 1" AND NOT #Cnv_Sensors."Pallet Detect 2" THEN
               #VTD_Control.Pallet_Loaded := 4; //Euro right alligned
               //Euro skewed to the right
           ELSIF #Cnv_Sensors."Pallet Detect 2" AND NOT #Cnv_Sensors."Pallet Detect 1" THEN
               #VTD_Control.Pallet_Loaded := 3; //Euro left alligned
               //Euro CENTERED
           ELSIF NOT #Cnv_Sensors."Pallet Detect 2" AND NOT #Cnv_Sensors."Pallet Detect 1" THEN
               #VTD_Control.Pallet_Loaded := 5;//'Euro';
               //Some unknown combination of sensors
           ELSE
               #VTD_Control.Pallet_Loaded := 1; //Unknown mythical pallet
           END_IF;

       ELSE
           //No Pallet
           #VTD_Control.Pallet_Loaded := 0; //No Pallet
       END_IF;

       // Locking pins state
       IF #LPL_Extended AND #LPR_Extended THEN
           #VTD_Control.LP_State := 1; //'Extended'
       ELSIF #LPL_Retracted AND #LPR_Retracted THEN
           #VTD_Control.LP_State := 2; //'Retracted'
       ELSE
           #VTD_Control.LP_State := 0; //'Unknown'
       END_IF;

       // Level detect
       #Level_Detect := #Level_Detect1 AND #Level_Detect2;

       //VTD extractor is docked
       IF #LPL_Extended AND #LPR_Extended AND #Level_Detect THEN

           #VTD_Control.Docked := TRUE;
       ELSE
           #VTD_Control.Docked := FALSE;
       END_IF;

       //Ultimate stop checks
       IF #Ulitmate_Creep AND #Ultimate_Slow AND #VTD_Control.Running THEN
           #VTD_Control.Motor_Speed := #VTD_Settings.Creep_Speed;
           #VTD_Control.Warning := 0; // Overtravel creep zone reached
       ELSIF NOT #Ulitmate_Creep AND #Ultimate_Slow AND #VTD_Control.Running THEN
           #VTD_Control.Motor_Speed := #VTD_Settings.Slow_Speed; // Overtravel creep zone reached
       END_IF;

       //Timeout of movement
       IF #VTD_Control.Mode = 2 OR #VTD_Control.Mode = 3 OR #VTD_Control.Mode = 4 THEN
           IF (#DestinationLevel - #CurrentlLevel = 1) AND #VTD_Control.Running THEN
               #Watchdog.TON(IN := TRUE,
                             PT := UINT_TO_TIME(#VTD_Settings.Transfer_Timeout_Up) * 1000);
           ELSIF (#DestinationLevel - #CurrentlLevel = 2) AND #VTD_Control.Running THEN
               #Watchdog.TON(IN := TRUE,
                             PT := UINT_TO_TIME(#VTD_Settings.Transfer_Timeout_Up) * 2000);
           ELSIF (#DestinationLevel - #CurrentlLevel = -1) AND #VTD_Control.Running THEN
               #Watchdog.TON(IN := TRUE,
                             PT := UINT_TO_TIME(#VTD_Settings.Transfer_Timeout_Down) * 1000);
           ELSIF (#DestinationLevel - #CurrentlLevel = -2) AND #VTD_Control.Running THEN
               #Watchdog.TON(IN := TRUE,
                             PT := UINT_TO_TIME(#VTD_Settings.Transfer_Timeout_Down) * 2000);
           ELSE
               #Watchdog.TON(IN := FALSE,
                             PT := T#0S);
           END_IF;
       END_IF;

       //Update Variables
       IF #VTD_Control.Current_Task_Type = 0 OR #VTD_Control.Current_Task_Type = 1 THEN
           #VTD_Control.SM_State := #State;
       ELSIF #VTD_Control.Current_Task_Type = 2 OR #VTD_Control.Current_Task_Type = 3 THEN
           #VTD_Control.SM_State := #I_State;
       END_IF;

       FOR #i := 1 TO "Settings_DB".System_Settings.Level_Count DO
           IF NOT "Control_DB".LCnv_Control[#i].Safety_Stop_Cnrl.Inputs.LP_Extended THEN
               #Cnvs1_NotExtended := true;
           END_IF;
           IF NOT "Control_DB".LCnv_Control[#i].Safety_Stop_Cnrl.Inputs.LP_Extended THEN
               #Cnvs2_NotExtended := true;
           END_IF;
       END_FOR;

       //Confirm whish level is below the extractor
       FOR #i := 0 TO "Settings_DB".System_Settings.Level_Count DO
           IF #VTD_Control.LE >= #VTD_Settings.Teach_Values.Levels_LE[#i] THEN
               #LevelBelowExtractor := #i;
           END_IF;
       END_FOR;

       #Stoppers_NotExtended := #Cnvs1_NotExtended (*AND #Cnvs2_NotExtended*);

       //AE ERROR
       IF "AE_Status_2".%X15 THEN
           #VTD_Control.AE_Error := 1;
       ELSE
           #VTD_Control.AE_Error := 0;
       END_IF;

       //Encoder Delta
       #VTD_Control.Encoder_Delta := ABS(#VTD_Control.AE - #VTD_Control.LE);

       //CURRENT LEVEL
       FOR #i := 0 TO #VTD_Settings.Highest_Level DO
           IF ABS(#VTD_Control.LE - #VTD_Settings.Teach_Values.Levels_LE[#i]) <= #VTD_Settings.VTD_Level_Granularity AND #Level_Detect THEN
               #VTD_Control.Current_Level := #i;
               EXIT;
           ELSE
               #VTD_Control.Current_Level := 99;
           END_IF;
       END_FOR;

       //Bypass linear encoder
       IF #VTD_Control.LE <> 0 THEN
           "LE_Bypass" := FALSE;
       END_IF;
   END_REGION

   REGION Auto/Semi-Auto Mode
           CASE #State OF
               0: //Idle
                   #DestinationLevel := #CurrentlLevel := 0;
                   "VTD_Move_To_Level_HMI_Tag" := 0;
                   IF (#VTD_Control.Mode = 3 AND #VTD_Control.Current_Task_Type = 1) OR #VTD_Control.Mode = 2 THEN
                       IF #VTD_Control.Instruction.Enable AND #VTD_Control.Error = 0 THEN
                           #VTD_Control.Enabled := TRUE;
                           #State := 10;
                       END_IF;
                   END_IF;

               10: //Standby
                   IF NOT #VTD_Control.Running AND #VTD_Control.Instruction.Move_To_Level <> 99 AND
                       ((#VTD_Control.Instruction.Task_ID > 0 OR #VTD_Control.Instruction.Task_Metadata <> '' AND #VTD_Control.Mode = 3 AND "Control_DB"."VTD_Order Table".Task_Type = 1) OR
                       (#VTD_Control.Mode = 2 AND #R_Execulte.Q))
                   THEN
                       IF #VTD_Control.Instruction.Move_To_Level = #VTD_Control.Current_Level AND #VTD_Control.Instruction.Move_To_Level <> 0 THEN
                           #VTD_Control.Warning := 1; //VTD already at level requested
                       //Go straght to the travel complete feedabck 
                       ELSIF (#VTD_Control.Shuttle_Loaded = 0 OR #VTD_Control.Shuttle_Loaded = 1) (*AND
                           (#VTD_Control.Pallet_Loaded = 0 OR #VTD_Control.Pallet_Loaded = 2 OR #VTD_Control.Pallet_Loaded = 3)*) THEN
                           #DestinationLevel := #VTD_Control.Instruction.Move_To_Level;
                           #CurrentlLevel := #VTD_Control.Current_Level;
                           #VTD_Control.Current_Task_ID := #VTD_Control.Instruction.Task_ID;
                           #State := 20;
                       // ELSIF #VTD_Control.Shuttle_Loaded = 2 THEN //24:11 Shuttle is not in the center of the extractor, to far forward
                       //     "Set_Bit_F"(Bit := 12,
                       //                 Bit_Value := 1,
                       //                 Var := #VTD_Control.VTD_Errors.Error_Word_2);
                       // ELSIF #VTD_Control.Shuttle_Loaded = 3 THEN //24:12 Shuttle is not in the center of the extractor, to far backward
                       //     "Set_Bit_F"(Bit := 13,
                       //                 Bit_Value := 1,
                       //                 Var := #VTD_Control.VTD_Errors.Error_Word_2);
                       // ELSIF #VTD_Control.Pallet_Loaded = 1 THEN //24:13 Pallet broken or not in position
                       //     "Set_Bit_F"(Bit := 14,
                       //                 Bit_Value := 1,
                       //                 Var := #VTD_Control.VTD_Errors.Error_Word_2);
                       // ELSE //24:14 Unknown load state
                       //     "Set_Bit_F"(Bit := 15,
                       //                 Bit_Value := 1,
                       //                 Var := #VTD_Control.VTD_Errors.Error_Word_2);
                       END_IF;

                   END_IF;

               20: //Extend all safety stoppers that are not in the up position
                   #VTD_Control.Running := TRUE;
                   #VTD_Control.Done := FALSE;// To report to order table
                   FOR #i := 1 TO "Settings_DB".System_Settings.Level_Count DO
                       IF NOT "Control_DB".LCnv_Control[#i].Safety_Stop_Cnrl.Inputs.LP_Extended THEN
                           "Control_DB".LCnv_Control[#i].Safety_Stop_Cnrl.Instruction.LP_Extend := TRUE;
                       END_IF;
                   END_FOR;
                   #State := 25;

               25: //Check to ensure the Safety stoppers are in the up position.    
                   FOR #i := 1 TO "Settings_DB".System_Settings.Level_Count DO
                       IF "Control_DB".LCnv_Control[#i].Safety_Stop_Cnrl.Inputs.LP_Extended THEN
                           "Control_DB".LCnv_Control[#i].Safety_Stop_Cnrl.Instruction.LP_Extend := FALSE;
                       END_IF;
                   END_FOR;
                   IF "Control_DB".LCnv_Control[1].Safety_Stop_Cnrl.Inputs.LP_Extended AND
                       "Control_DB".LCnv_Control[2].Safety_Stop_Cnrl.Inputs.LP_Extended AND
                       "Control_DB".LCnv_Control[3].Safety_Stop_Cnrl.Inputs.LP_Extended THEN
                       #State := 30;
                   END_IF;

               30: //Undock the VTD
                   IF #VTD_Control.Docked OR (#VTD_Control.LE < #VTD_Settings.Teach_Values.Levels_LE[#LevelBelowExtractor]+ 50 AND
                       #VTD_Control.LE > #VTD_Settings.Teach_Values.Levels_LE[#LevelBelowExtractor]) THEN
                       IF #VTD_Control.LP_State = 1 THEN //extended
                           #VTD_Control.Motor_Speed := #VTD_Settings.Dock_speed;
                           #VTD_Control.Motor_UP := TRUE;
                           #Position_Offset := #VTD_Control.LE + 40;
                           #State := 35;
                       ELSIF #VTD_Control.LP_State = 2 THEN //retracted
                           #State := 45;
                       ELSE //24:4 Docking pins in an known state
                           "Set_Bit_F"(Bit := 5,
                                       Bit_Value := 1,
                                       Var := #VTD_Control.VTD_Errors.Error_Word_2);
                       END_IF;
                   ELSE
                       #Position_Offset := #VTD_Control.LE - 5;
                       #State := 35;
                   END_IF;

               35: //Retract the docking pins
                   IF NOT #Level_Detect AND #VTD_Control.LE >= #Position_Offset THEN //change back to the original condition
                       #VTD_Control.Motor_Speed := 0;
                       #VTD_Control.Motor_UP := FALSE;
                       #LPR_Retract := #LPL_Retract := TRUE;
                       #LP_Timer(IN := TRUE,
                                 PT := UINT_TO_TIME(#VTD_Settings.Lockpins_Timeout_Retract));

                       IF #LPR_Retracted THEN
                           #LPR_Retract := FALSE;
                       END_IF;
                       IF #VTD_Control.Inputs.LPL_Retracted THEN
                           #LPL_Retract := FALSE;
                       END_IF;

                       IF #VTD_Control.LP_State = 2 THEN
                           #State := 40;
                       END_IF;
                   END_IF;

               40: //Check docking pins have been retracted
                   IF #VTD_Control.LP_State = 2 THEN
                       #LP_Timer(IN := FALSE,
                                 PT := T#0S);
                       #LPR_Retract := #LPL_Retract := FALSE;
                       #State := 45;
                   END_IF;

               45: //Start moving towards the level required
                   //Check load type and set extractor speed
                   IF #VTD_Control.Shuttle_Loaded = 0 AND #VTD_Control.Pallet_Loaded = 0 THEN 
                       #VTD_Control.Motor_Speed := #VTD_Settings.Empty_Speed;
                   ELSIF #VTD_Control.Shuttle_Loaded = 1 AND #VTD_Control.Pallet_Loaded = 0 THEN
                       #VTD_Control.Motor_Speed := #VTD_Settings.Shuttle_Speed;
                   ELSIF #VTD_Control.Shuttle_Loaded = 0 AND (#VTD_Control.Pallet_Loaded > 0) THEN
                       #VTD_Control.Motor_Speed := #VTD_Settings.Pallet_Speed;
                   ELSIF #VTD_Control.Shuttle_Loaded = 1 AND (#VTD_Control.Pallet_Loaded > 0) THEN
                       #VTD_Control.Motor_Speed := #VTD_Settings.Loaded_Speed;
                   END_IF;

                   #DestPosition := #VTD_Settings.Teach_Values.Levels_LE[#VTD_Control.Instruction.Move_To_Level];
                   #SetUpSpeed := #VTD_Control.Motor_Speed;

                   //VTD needs to move up
                   IF #VTD_Control.LE < #DestPosition THEN
                       #VTD_Control.Motor_UP := TRUE;
                       #State := 50;
                       //VTD needs to move down
                   ELSIF #VTD_Control.LE > #DestPosition THEN
                       #VTD_Control.Motor_Down := TRUE;
                       #State := 65; //change to 65
                   END_IF;

               50: //travel upwards to designated level
                   #ChangeToLow[1] := ABS((#VTD_Settings.Slowdown_Count_LE / 100) * 80); (* 80% *) //80  600mm
                   #ChangeToLow[2] := ABS((#VTD_Settings.Slowdown_Count_LE / 100) * 60); (* 60% *) //60
                   #ChangeToLow[3] := ABS((#VTD_Settings.Slowdown_Count_LE / 100) * 40); (* 40% *) //40
                   #ChangeToLow[4] := ABS((#VTD_Settings.Slowdown_Count_LE / 100) * 20); (* 20% *) //20 60

                   //switch to fast freq Low UP
                   IF ABS(#DestPosition - #VTD_Control.LE) > #VTD_Settings.Slowdown_Count_LE THEN
                       #VTD_Control.Motor_Speed := #SetUpSpeed; //5
                       //switch to low freq
                   ELSIF ABS(#DestPosition - #VTD_Control.LE) <= #VTD_Settings.Slowdown_Count_LE
                       AND ABS(#DestPosition - #VTD_Control.LE) > #ChangeToLow[1] THEN
                       #VTD_Control.Motor_Speed := #VTD_Settings.Slow_Calib_Speed * 1.8; //5 * 1.8 = 9%
                   ELSIF ABS(#DestPosition - #VTD_Control.LE) <= #ChangeToLow[1]
                       AND ABS(#DestPosition - #VTD_Control.LE) > #ChangeToLow[2] THEN
                       #VTD_Control.Motor_Speed := #VTD_Settings.Slow_Calib_Speed * 1.6; //5 * 1.6 = 8%
                   ELSIF ABS(#DestPosition - #VTD_Control.LE) <= #ChangeToLow[2]
                       AND ABS(#DestPosition - #VTD_Control.LE) > #ChangeToLow[3] THEN
                       #VTD_Control.Motor_Speed := #VTD_Settings.Slow_Calib_Speed * 1.4; //5 * 1.4 = 7%
                   ELSIF ABS(#DestPosition - #VTD_Control.LE) <= #ChangeToLow[3]
                       AND ABS(#DestPosition - #VTD_Control.LE) > #ChangeToLow[4] THEN
                       #VTD_Control.Motor_Speed := #VTD_Settings.Slow_Calib_Speed * 1.2; //5 * 1.2 = 6%
                   ELSIF ABS(#DestPosition - #VTD_Control.LE) <= #ChangeToLow[4] THEN
                       #VTD_Control.Motor_Speed := #VTD_Settings.Slow_Calib_Speed; //5%
                       #State := 55;
                   END_IF;

               55: // Travel upwards using slow speed towards required floor
                   IF #VTD_Control.LE > #VTD_Settings.Teach_Values.Levels_LE[#VTD_Control.Instruction.Move_To_Level] - #VTD_Settings.Creep_Count_LE
                   THEN
                       #VTD_Control.Motor_Speed := #VTD_Settings.Creep_Speed; //3% - 60mm 
                       #State := 60;
                   END_IF;

               60: // Travel past the level in order to extend the docking pins
                   IF #VTD_Control.LE > #VTD_Settings.Teach_Values.Levels_LE[#VTD_Control.Instruction.Move_To_Level] + #VTD_Settings.Creep_Count_LE
                   THEN
                       #VTD_Control.Motor_Speed := 0;
                       #VTD_Control.Motor_UP := FALSE;
                       #State := 80;
                   END_IF;

               65: //travel Downwards to designated level   
                   #ChangeToLow[1] := ABS((#VTD_Settings.Slowdown_Count_LE / 100) * 80); (* 80% *) //80
                   #ChangeToLow[2] := ABS((#VTD_Settings.Slowdown_Count_LE / 100) * 60); (* 60% *) //60
                   #ChangeToLow[3] := ABS((#VTD_Settings.Slowdown_Count_LE / 100) * 40); (* 40% *) //40
                   #ChangeToLow[4] := ABS((#VTD_Settings.Slowdown_Count_LE / 100) * 20); (* 20% *) //20
                   //switch to fast freq Low UP
                   IF ABS(#DestPosition - #VTD_Control.LE) > #VTD_Settings.Slowdown_Count_LE THEN
                       #VTD_Control.Motor_Speed := #SetUpSpeed;
                       //switch to low freq
                   ELSIF ABS(#DestPosition - #VTD_Control.LE) <= #VTD_Settings.Slowdown_Count_LE
                       AND ABS(#DestPosition - #VTD_Control.LE) > #ChangeToLow[1] THEN
                       #VTD_Control.Motor_Speed := #VTD_Settings.Slow_Calib_Speed * 1.8;
                   ELSIF ABS(#DestPosition - #VTD_Control.LE) <= #ChangeToLow[1]
                       AND ABS(#DestPosition - #VTD_Control.LE) > #ChangeToLow[2] THEN
                       #VTD_Control.Motor_Speed := #VTD_Settings.Slow_Calib_Speed * 1.6;
                   ELSIF ABS(#DestPosition - #VTD_Control.LE) <= #ChangeToLow[2]
                       AND ABS(#DestPosition - #VTD_Control.LE) > #ChangeToLow[3] THEN
                       #VTD_Control.Motor_Speed := #VTD_Settings.Slow_Calib_Speed * 1.4;
                   ELSIF ABS(#DestPosition - #VTD_Control.LE) <= #ChangeToLow[3]
                       AND ABS(#DestPosition - #VTD_Control.LE) > #ChangeToLow[4] THEN
                       #VTD_Control.Motor_Speed := #VTD_Settings.Slow_Calib_Speed * 1.2;
                   ELSIF ABS(#DestPosition - #VTD_Control.LE) <= #ChangeToLow[4] THEN
                       #VTD_Control.Motor_Speed := #VTD_Settings.Slow_Calib_Speed;
                       #State := 70;
                   END_IF;

               70: // Travel downwards using slow speed towards required floor 
                   IF #VTD_Control.LE < #VTD_Settings.Teach_Values.Levels_LE[#VTD_Control.Instruction.Move_To_Level] + #VTD_Settings.Creep_Count_LE
                   THEN
                       #VTD_Control.Motor_Speed := 0;
                       #VTD_Control.Motor_Down := FALSE;
                       #State := 80;
                   END_IF;

               80: //Extend Docking pins
                   IF #VTD_Control.LP_State = 2 AND NOT #Level_Detect THEN 
                       #LPL_Extend := #LPR_Extend := TRUE;
                       #LP_Timer(IN := TRUE,
                                 PT := UINT_TO_TIME(#VTD_Settings.Lockpins_Timeout_Extend));
                   ELSIF #VTD_Control.LP_State <> 1 AND NOT #Level_Detect THEN 
                       #LPL_Extend := #LPR_Extend := TRUE;
                   ELSIF #VTD_Control.LP_State = 1 THEN
                       #State := 85;
                   END_IF;


               85: // Wait for docking pins to extend
                   IF #VTD_Control.LP_State = 1 AND NOT #Level_Detect THEN
                       #LP_Timer(IN := FALSE,
                                 PT := T#0S);
                       #LPL_Extend := #LPR_Extend := FALSE;
                       #VTD_Control.Motor_Speed := #VTD_Settings.Dock_speed;
                       #VTD_Control.Motor_Down := TRUE;
                       #State := 90;
                   END_IF;

               90: // Dock the VTD
                   //Using the Linear Encoder for comparation and Release tension in the VTD chain
                   IF ABS(#VTD_Control.LE - #DestPosition) <= (#VTD_Settings.Level_Detect_LE) AND NOT #CS_TImer.Q THEN
                       #CS_TImer(IN := TRUE,
                                 PT := UINT_TO_TIME(#VTD_Settings.Chain_Slack_Timeout));
                   END_IF;
                   IF #CS_TImer.Q THEN
                       #VTD_Control.Motor_Speed := 0;
                       #VTD_Control.Motor_Down := FALSE;
                       #CS_TImer(IN := FALSE,
                                 PT := T#0S);
                       #State := 95;
                   END_IF;

               95: // Dock the VTD
                   //Check the level detect sensors
                   IF (#Level_Detect1 AND NOT #Level_Detect2) OR
                       (NOT #Level_Detect1 AND #Level_Detect2) THEN
                       #LD_Timer(IN := TRUE,
                                 PT := UINT_TO_TIME(#VTD_Settings.Level_Detect_Timeout));
                   ELSE
                       #LD_Timer(IN := FALSE,
                                 PT := T#0s);
                   END_IF;

                       IF #Level_Detect THEN
                           #Watchdog(IN := FALSE,
                                     PT := T#0S);
                           #State := 100;
                       END_IF;

               100: //Wait for Movement completion ack  
                   //Reset timers
                   #LP_Timer(IN := FALSE,
                             PT := T#0s);
                   #Watchdog(IN := FALSE,
                             PT := T#0s);
                   #LD_Timer(IN := FALSE,
                             PT := T#0s);
                   #CS_TImer(IN := FALSE,
                             PT := T#0s);

                   #VTD_Control.Motor_Speed := 0;
                   IF #VTD_Control.Mode = 3 THEN //VTD in Auto

                       IF "Control_DB"."VTD_Order Table".Movement_Request_Complete_Ack THEN
                           #VTD_Control.Current_Task_ID := 0;
                           #VTD_Control.Running := FALSE;
                           #VTD_Control.Done := TRUE;// To report to order table
                           #State := 0;
                           // "Control_DB".WMS_OPC_UA.Movement_Request_Complete_Ack := FALSE;
                       END_IF;
                   ELSIF #VTD_Control.Mode = 2 THEN //VTD in Semi-Auto
                       #VTD_Control.Current_Task_ID := 0;
                       "VTD_Move_To_Level_HMI_Tag" := 0;
                       #VTD_Control.Running := FALSE;
                       #State := 0;
                   END_IF;

               400: // Error state
                   #VTD_Control.Done := FALSE;// To report to order table
                   #VTD_Control.Motor.Enable := FALSE;
                   #VTD_Control.Motor_UP := FALSE;
                   #VTD_Control.Motor_Down := FALSE;
                   #VTD_Control.Running := FALSE;
                   #VTD_Control.Stopped := TRUE;
                   #VTD_Control.Motor.Speed := 0;
                   #VTD_Control.Motor.Forward := FALSE;
                   #VTD_Control.Motor.Reverse := FALSE;
                   #LPL_Extend := #LPR_Extend := FALSE;
                   #LPL_Retract := #LPR_Retract := FALSE;
                   //Reset timers
                   #LP_Timer(IN := FALSE,
                             PT := T#0s);
                   #Watchdog(IN := FALSE,
                             PT := T#0s);
                   #LD_Timer(IN := FALSE,
                             PT := T#0s);
                   #CS_TImer(IN := FALSE,
                             PT := T#0s);
                   IF #VTD_Control.Instruction.Reset THEN
                       #VTD_Control.Instruction.Move_To_Level := 0;
                       "VTD_Move_To_Level_HMI_Tag" := 0;
                       #VTD_Control.Error := FALSE;
                       #VTD_Control.Warning := 0;
                       #VTD_Control.Stopped := FALSE;
                       #VTD_Control.Current_Task_Type := 0;
                       #VTD_Control.VTD_Errors.Error_Word_1 := 0;
                       #VTD_Control.VTD_Errors.Error_Word_2 := 0;
                       #VTD_Control.VTD_Errors.Error_Word_3 := 0;
                       #VTD_Control.VTD_Errors.Error_Word_4 := 0;
                       #State := 0;
                   END_IF;

               500: //MANUAL MODE
                   IF #VTD_Control.Error = 0 THEN

                       //VTD
                       IF #VTD_Control.Instruction.Manual_Up AND NOT "Upper Ultimate" THEN
                           #VTD_Control.Motor_UP := TRUE;
                           #VTD_Control.Running := TRUE;
                           IF NOT (#Ultimate_Slow OR #Ulitmate_Creep) THEN
                               #VTD_Control.Motor_Speed := #VTD_Settings.Manual_Speed;
                           END_IF;
                       ELSIF #VTD_Control.Instruction.Manual_Down AND NOT "Lower Ultimate" THEN
                           #VTD_Control.Motor_Down := TRUE;
                           #VTD_Control.Running := TRUE;
                           IF NOT (#Ultimate_Slow OR #Ulitmate_Creep) THEN
                               #VTD_Control.Motor_Speed := #VTD_Settings.Manual_Speed;
                           END_IF;
                       ELSE
                           #VTD_Control.Motor_Speed := 0;
                           #VTD_Control.Running := FALSE;
                           #VTD_Control.Motor_Down := FALSE;
                           #VTD_Control.Motor_UP := FALSE;
                       END_IF;

                       //LOCKING PINS RIGHT 
                       IF NOT #VTD_Control.Running AND #VTD_Control.Instruction.Manual_LP_Extend
                           AND NOT #LPR_Extended THEN
                           #LPR_Extend := TRUE;
                       ELSIF NOT #VTD_Control.Running AND #VTD_Control.Instruction.Manual_LP_Retract
                           AND NOT #LPR_Retracted THEN
                           #LPR_Retract := TRUE;
                       ELSE
                           #LPR_Extend := FALSE;
                           #LPR_Retract := FALSE;
                       END_IF;

                       //LOCKING PINS LEFT 
                       IF NOT #VTD_Control.Running AND #VTD_Control.Instruction.Manual_LP_Extend
                           AND NOT #LPL_Extended THEN
                           #LPL_Extend := TRUE;
                       ELSIF NOT #VTD_Control.Running AND #VTD_Control.Instruction.Manual_LP_Retract
                           AND NOT #LPL_Retracted THEN
                           #LPL_Retract := TRUE;
                       ELSE
                           #LPL_Extend := FALSE;
                           #LPL_Retract := FALSE;
                       END_IF;

                       IF #VTD_Control.Mode <> 1 AND #VTD_Control.Mode <> 5 THEN
                           #State := 0;
                       END_IF;

                       IF #LPR_Extend OR #LPL_Extend THEN
                           #LP_Timer(IN := TRUE,
                                     PT := UINT_TO_TIME(#VTD_Settings.Lockpins_Timeout_Extend));
                       ELSIF #LPR_Retract OR #LPL_Retract THEN
                           #LP_Timer(IN := TRUE,
                                     PT := UINT_TO_TIME(#VTD_Settings.Lockpins_Timeout_Retract));
                       ELSE
                           #LP_Timer(IN := FALSE,
                                     PT := T#0S);
                       END_IF;
                   END_IF;
           END_CASE;
   END_REGION

   REGION Shuttle Interlock
       // VTD needs to be in Auto mode to perform a Shuttle interlock
       CASE #I_State OF
           0:
               IF #VTD_Control.Mode = 3 AND #VTD_Control.Shuttle_Interlock.Interlock_Request AND #VTD_Control.Shuttle_Interlock.Shuttle_Interlock_Task_ID > 0 THEN
                   #I_State := 10;
               END_IF;

               10: //Standby

                   //Start by decoding all the IDs of the devices pertaining to the VTD in question on that level
                   "ID_Decode_F"(ID := #VTD_Settings.ID,
                                 ID_Decoded := #VTD_ID_Decoded);
                   "ID_Decode_F"(ID := "Settings_DB".LCnv_Settings[#VTD_Control.Current_Level].ID,
                                 ID_Decoded := #Cnv_ID_Decoded);

                   // Ensure the VTD is in a state that it can perform an interlock
                   IF #VTD_Control.Docked AND NOT #VTD_Control.Running AND (#VTD_Control.Shuttle_Loaded = 0 OR #VTD_Control.Shuttle_Loaded = 1) AND #VTD_Control.Error = 0 THEN
                       // Check to make sure the VTD and Shuttle are not both loaded
                       IF #VTD_Control.Pallet_Loaded = 1 THEN
                           #VTD_Control.Warning := 1; // Both the VTD and Shuttles are loaded, can't perform the interlock
                       ELSE
                           //Check that shuttle is on the correct floor, that the start location given and the shuttle actual position matches and the destination is the correct extractor barcode
                           IF (*#VTD_Control.Current_Level = "Shuttle_MQTT_DB".Shuttle_MQTT[#VTD_Control.Shuttle_Interlock.Shuttle_ID].Message.Shuttle_Status.Floor
                               AND*) #VTD_Control.Shuttle_Interlock.Shuttle_Start_Location = "Shuttle_MQTT_DB".Shuttle_MQTT[#VTD_Control.Shuttle_Interlock.Shuttle_ID].Message.Shuttle_Status.Position_ID
                               (*AND "Shuttle_MQTT_DB".Shuttle_MQTT[#VTD_Control.Shuttle_Interlock.Shuttle_ID].Message.Shuttle_Status.Destination_ID = "Settings_DB".ECnv_Settings.Barcode_ID*)THEN

                               //Check in which Buffer conveyor the shuttle is located
                               IF "Settings_DB".LCnv_Settings[#VTD_Control.Current_Level].Barcode_ID =
                                   #VTD_Control.Shuttle_Interlock.Shuttle_Start_Location THEN
                                   #VTD_Control.Running := TRUE;
                                   #I_State := 20;
                               ELSIF "Settings_DB".ECnv_Settings.Barcode_ID =
                                   #VTD_Control.Shuttle_Interlock.Shuttle_Start_Location AND
                                   "Control_DB"."VTD_Order Table".Destination_Location = "Settings_DB".LCnv_Settings[#VTD_Control.Current_Level].Barcode_ID THEN
                                   #VTD_Control.Running := TRUE;
                                   #I_State := 20;
                               ELSE
                                   #VTD_Control.Warning := 2; // Shuttle interlock start location not buffer conveyor of VTD
                               END_IF;
                           ELSE
                               #VTD_Control.Warning := 3; // Cant interlock as shuttle and VTD level mismatch
                           END_IF;
                       END_IF;
                   ELSE
                       #VTD_Control.Warning := 4; // VTD not ready for interlock 
                   END_IF;


               20: //Drop safety stops
                   IF #Cnv_ID_Decoded.Level = #VTD_Control.Current_Level THEN
                       "Control_DB".LCnv_Control[#VTD_Control.Current_Level].Safety_Stop_Cnrl.Instruction.LP_Retract := TRUE;
                       #I_State := 30;
                   ELSE
                       #VTD_Control.Error := TRUE; //24:16 Cannot find the correct safety pins to drop.
                       "Set_Bit_F"(Bit := 1,
                                   Bit_Value := 1,
                                   Var := #VTD_Control.VTD_Errors.Error_Word_3);
                       // #I_State := 400;
                   END_IF;

               //////////////////////////////////////////////////////////////////////////////////////////////////////////////////////////////////////////////////////////////////    
               30: //Confirm safety stops are down at the correct location
                   //Send ready to interlock
                   IF "Control_DB".LCnv_Control[#VTD_Control.Current_Level].Safety_Stop_Cnrl.LP_State = 0 THEN //RETRACTED
                       "Control_DB".LCnv_Control[#VTD_Control.Current_Level].Safety_Stop_Cnrl.Instruction.LP_Retract := FALSE;
                       #VTD_Control.Shuttle_Interlock.Ready_To_Interlock := TRUE;
                       #I_State := 40;
                   END_IF;

               ////////////////////////////////////////////////////////////////////////////////////////////////////////////////////////////////////////////////////////////////////
               40: //Wait for shuttle to move in or out VTD
                   //Add timer for shuttle transfer to occur
                   IF "Control_DB"."VTD_Order Table".Destination_Location = "Settings_DB".ECnv_Settings.Barcode_ID THEN
                       IF "Settings_DB".ECnv_Settings.Barcode_ID = "Shuttle_MQTT_DB".Shuttle_MQTT[#VTD_Control.Shuttle_Interlock.Shuttle_ID].Message.Shuttle_Status.Position_ID
                           AND "Shuttle_MQTT_DB".Shuttle_MQTT[#VTD_Control.Shuttle_Interlock.Shuttle_ID].Message.Shuttle_Status.Operational_State = 'IDLE' THEN
                           "Control_DB".LCnv_Control[#VTD_Control.Current_Level].Safety_Stop_Cnrl.Instruction.LP_Extend := TRUE;
                           #I_State := 50;
                       END_IF;
                   ELSIF "Control_DB"."VTD_Order Table".Destination_Location = "Settings_DB".LCnv_Settings[#VTD_Control.Current_Level].Barcode_ID THEN
                       IF "Settings_DB".LCnv_Settings[#VTD_Control.Current_Level].Barcode_ID = "Shuttle_MQTT_DB".Shuttle_MQTT[#VTD_Control.Shuttle_Interlock.Shuttle_ID].Message.Shuttle_Status.Position_ID
                           AND "Shuttle_MQTT_DB".Shuttle_MQTT[#VTD_Control.Shuttle_Interlock.Shuttle_ID].Message.Shuttle_Status.Operational_State = 'IDLE' THEN
                           "Control_DB".LCnv_Control[#VTD_Control.Current_Level].Safety_Stop_Cnrl.Instruction.LP_Extend := TRUE;
                           #I_State := 50;
                       END_IF;
                   END_IF;

               //////////////////////////////////////////////////////////////////////////////////////////////////////////////////////////////////////////////////////////////////////////  
               50: //Check own sensors for shuttle/pallet state
                   #IEC_Timer_0_Instance_1(IN:=TRUE,
                                           PT:=T#5S);
                   IF "Control_DB".LCnv_Control[#VTD_Control.Current_Level].Safety_Stop_Cnrl.LP_State = 1 //EXTENDED
                       AND "Control_DB".ECnv_Control.Shuttle_In_Place THEN
                       "Control_DB".LCnv_Control[#VTD_Control.Current_Level].Safety_Stop_Cnrl.Instruction.LP_Extend := FALSE;
                       #VTD_Control.Shuttle_Interlock.Interlock_Complete := TRUE;
                       #I_State := 60;
                   ELSIF #IEC_Timer_0_Instance_1.Q THEN
                       #VTD_Control.Error := TRUE; //24:17 Error occured during interlock final check
                       "Set_Bit_F"(Bit := 2,
                                   Bit_Value := 1,
                                   Var := #VTD_Control.VTD_Errors.Error_Word_3);
                       #I_State := 400;
                   END_IF;

               60://Clear Vars
                   #IEC_Timer_0_Instance_1(IN := FALSE,
                                           PT := T#0s);
                   #IEC_Timer_0_Instance_2(IN := FALSE,
                                           PT := T#0s);
                   IF #VTD_Control.Shuttle_Interlock.Interlock_Complete_Ack THEN
                       #VTD_Control.Shuttle_Interlock.Ready_To_Interlock := FALSE;
                       #VTD_Control.Shuttle_Interlock.Interlock_Complete := FALSE;
                       #VTD_Control.Running := FALSE;
                       #I_State := 0;
                   END_IF;

               400://ERROR MODE
                   #IEC_Timer_0_Instance_1(IN := FALSE,
                                           PT := T#0s);
                   #IEC_Timer_0_Instance_2(IN := FALSE,
                                           PT := T#0s);
                   #Interlock_Timer(IN := FALSE,
                                    PT := T#0s);
                   #VTD_Control.Running := FALSE;
                   #VTD_Control.Shuttle_Interlock.Interlock_Complete := FALSE;
                   #VTD_Control.Shuttle_Interlock.Ready_To_Interlock := FALSE;
                   "Control_DB".LCnv_Control[#VTD_Control.Current_Level].Safety_Stop_Cnrl.Instruction.LP_Extend := FALSE;
                   "Control_DB".LCnv_Control[#VTD_Control.Current_Level].Safety_Stop_Cnrl.Instruction.LP_Extend := FALSE;
                   "Control_DB".LCnv_Control[#VTD_Control.Current_Level].Safety_Stop_Cnrl.Instruction.LP_Retract := FALSE;
                   "Control_DB".LCnv_Control[#VTD_Control.Current_Level].Safety_Stop_Cnrl.Instruction.LP_Retract := FALSE;
                   IF #VTD_Control.Instruction.Reset THEN
                       #VTD_Control.VTD_Errors.Error_Word_3 := 0;
                       #I_State := 0;
                   END_IF;
               END_CASE;
           #Interlock_Timer(IN := #I_State >= 40 AND #I_State <= 50,
                            PT := UINT_TO_TIME("Settings_DB".System_Settings.Shuttle_Interlock_Timeout) * 1000);

   END_REGION

   REGION Cyclic Error Checks
       IF NOT "Main_Safety_RTG1_DB".SAFETY_OK_VTD THEN //21:1
           "Set_Bit_F"(Bit := 0,
                       Bit_Value := 1,
                       Var := #VTD_Control.VTD_Errors.Error_Word_1);
       END_IF;

       IF "VTD_Stop_HMI_Tag" THEN //21:2
           "Set_Bit_F"(Bit := 1,
                       Bit_Value := 1,
                       Var := #VTD_Control.VTD_Errors.Error_Word_1);
       END_IF;

       IF NOT "Overtravel Upper Limit - CH1" THEN //21:3
           "Set_Bit_F"(Bit := 2,
                       Bit_Value := 1,
                       Var := #VTD_Control.VTD_Errors.Error_Word_1);
       END_IF;

       IF NOT "Overtravel Lower Limit - CH1" THEN //21:4
           "Set_Bit_F"(Bit := 3,
                       Bit_Value := 1,
                       Var := #VTD_Control.VTD_Errors.Error_Word_1);
       END_IF;

       IF (#VTD_Control.Mode = 1 OR #VTD_Control.Mode = 5) AND #VTD_Control.Instruction.Manual_Up AND
           #VTD_Control.LE > #VTD_Settings.Teach_Values.Levels_LE[#VTD_Settings.Highest_Level] + #VTD_Settings.Creep_Count_LE THEN //21:5
           "Set_Bit_F"(Bit := 4,
                       Bit_Value := 1,
                       Var := #VTD_Control.VTD_Errors.Error_Word_1);
       END_IF;

       "R_TRIG_DB_3"(CLK:=#VTD_Control.Mode = 3);

       IF NOT #VTD_Control.Docked AND "R_TRIG_DB_3".Q THEN //22:1
           "Set_Bit_F"(Bit := 8,
                       Bit_Value := 1,
                       Var := #VTD_Control.VTD_Errors.Error_Word_1);
       END_IF;

       IF NOT #Level_Detect AND "R_TRIG_DB_3".Q THEN //22:2
           "Set_Bit_F"(Bit := 9,
                       Bit_Value := 1,
                       Var := #VTD_Control.VTD_Errors.Error_Word_1);
       END_IF;

       // IF "R_TRIG_DB_3".Q AND NOT ((#VTD_Control.LE < #VTD_Settings.Teach_Values.Levels_LE[1] + #VTD_Settings.VTD_Level_Granularity
       //     AND #VTD_Control.LE > #VTD_Settings.Teach_Values.Levels_LE[1] - #VTD_Settings.VTD_Level_Granularity)
       //     OR
       //     (#VTD_Control.LE < #VTD_Settings.Teach_Values.Levels_LE[2] + #VTD_Settings.VTD_Level_Granularity
       //     AND #VTD_Control.LE > #VTD_Settings.Teach_Values.Levels_LE[2] - #VTD_Settings.VTD_Level_Granularity)
       //     OR
       //     (#VTD_Control.LE < #VTD_Settings.Teach_Values.Levels_LE[3] + #VTD_Settings.VTD_Level_Granularity
       //     AND #VTD_Control.LE > #VTD_Settings.Teach_Values.Levels_LE[3] - #VTD_Settings.VTD_Level_Granularity))
       // THEN //22:3
       //         "Set_Bit_F"(Bit := 10,
       //                     Bit_Value := 1,
       //                     Var := #VTD_Control.VTD_Errors.Error_Word_1);
       // END_IF;

       IF #VTD_Control.Docked AND (#LPL_Retract OR #LPR_Retract) THEN //22:5
           "Set_Bit_F"(Bit := 12,
                       Bit_Value := 1,
                       Var := #VTD_Control.VTD_Errors.Error_Word_1);
       END_IF;

       #IEC_Timer_0_Instance(IN := #VTD_Control.LE <= (#VTD_Settings.Teach_Values.Levels_LE[#LevelBelowExtractor] + 1) AND #VTD_Control.Instruction.Manual_Down,
                             PT := t#300ms);

       //LINEAR ENCODER ERROR
       "IEC_Timer_0_DB_8".TON(IN := "LE_Status".%X0 OR "LE_Status".%X1 OR
                              #VTD_Control.LE < #VTD_Settings.VTD_Min_Height OR
                              #VTD_Control.LE > #VTD_Settings.VTD_Max_Heigh,
                              PT := t#500ms);
       IF NOT "LE_Bypass" AND "IEC_Timer_0_DB_8".Q THEN
           "Set_Bit_F"(Bit := 4,
                       Bit_Value := 1,
                       Var := #VTD_Control.VTD_Errors.Error_Word_3);
           "IEC_Timer_0_DB_8".TON (IN := FALSE,
                                   PT := T#0s);
       END_IF;

